(* IEC 61131-3 sources: BioPrint-Automation-Suite/projects/02_bioprint_pid/plc/src, 4 files *)

(* ---- DUT_ReferenceVectors.st ---- *)
(* =============================================================================
   DUT_ReferenceVectors — GENERATED by plc/generate_test_vectors.py. Do not edit.
   Struct types for GVL_ReferenceVectors (two DUTs in TwinCAT / CODESYS).
   ============================================================================= *)
TYPE ST_PidVector :
STRUCT
    lrSetpoint    : LREAL;
    lrMeasurement : LREAL;
    lrOutput      : LREAL;
    lrITerm       : LREAL;
END_STRUCT
END_TYPE

TYPE ST_WestgardVector :
STRUCT
    diStep     : DINT;
    lrValue    : LREAL;
    bWarn12s   : BOOL;
    bReject13s : BOOL;
    bReject22s : BOOL;
END_STRUCT
END_TYPE

(* ---- GVL_ReferenceVectors.st ---- *)
(* =============================================================================
   GVL_ReferenceVectors — GENERATED by plc/generate_test_vectors.py. Do not edit.
   Inputs and outputs of the Python reference implementation for the default
   scenario (config/default.toml), replayed scan by scan in the TcUnit tests.
   Types: DUT_ReferenceVectors.st
   ============================================================================= *)
{attribute 'qualified_only'}
VAR_GLOBAL CONSTANT
    N_VECTORS       : INT   := 300;
    LR_BASELINE_SD  : LREAL := 2.918663164239998E-01;
    aPid : ARRAY[1..300] OF ST_PidVector := [
        (lrSetpoint := 2.300000000000000E+02, lrMeasurement := 2.504570756196317E+01, lrOutput := 1.000000000000000E+02, lrITerm := 0.000000000000000E+00),
        (lrSetpoint := 2.300000000000000E+02, lrMeasurement := 2.559400238406393E+01, lrOutput := 1.000000000000000E+02, lrITerm := 0.000000000000000E+00),
        (lrSetpoint := 2.300000000000000E+02, lrMeasurement := 2.721106767937097E+01, lrOutput := 1.000000000000000E+02, lrITerm := 0.000000000000000E+00),
        (lrSetpoint := 2.300000000000000E+02, lrMeasurement := 2.906538770745868E+01, lrOutput := 1.000000000000000E+02, lrITerm := 0.000000000000000E+00),
        (lrSetpoint := 2.300000000000000E+02, lrMeasurement := 3.083779911570193E+01, lrOutput := 1.000000000000000E+02, lrITerm := 0.000000000000000E+00),
        (lrSetpoint := 2.300000000000000E+02, lrMeasurement := 3.344406655918265E+01, lrOutput := 1.000000000000000E+02, lrITerm := 0.000000000000000E+00),
        (lrSetpoint := 2.300000000000000E+02, lrMeasurement := 3.640825075871666E+01, lrOutput := 1.000000000000000E+02, lrITerm := 0.000000000000000E+00),
        (lrSetpoint := 2.300000000000000E+02, lrMeasurement := 3.928242815999355E+01, lrOutput := 1.000000000000000E+02, lrITerm := 0.000000000000000E+00),
        (lrSetpoint := 2.300000000000000E+02, lrMeasurement := 4.241953904612176E+01, lrOutput := 1.000000000000000E+02, lrITerm := 0.000000000000000E+00),
        (lrSetpoint := 2.300000000000000E+02, lrMeasurement := 4.550594203217187E+01, lrOutput := 1.000000000000000E+02, lrITerm := 0.000000000000000E+00),
        (lrSetpoint := 2.300000000000000E+02, lrMeasurement := 4.907188733629471E+01, lrOutput := 1.000000000000000E+02, lrITerm := 0.000000000000000E+00),
        (lrSetpoint := 2.300000000000000E+02, lrMeasurement := 5.243664392789950E+01, lrOutput := 1.000000000000000E+02, lrITerm := 0.000000000000000E+00),
        (lrSetpoint := 2.300000000000000E+02, lrMeasurement := 5.576754175418417E+01, lrOutput := 1.000000000000000E+02, lrITerm := 0.000000000000000E+00),
        (lrSetpoint := 2.300000000000000E+02, lrMeasurement := 5.940904962608809E+01, lrOutput := 1.000000000000000E+02, lrITerm := 0.000000000000000E+00),
        (lrSetpoint := 2.300000000000000E+02, lrMeasurement := 6.282668317532421E+01, lrOutput := 1.000000000000000E+02, lrITerm := 0.000000000000000E+00),
        (lrSetpoint := 2.300000000000000E+02, lrMeasurement := 6.617020839567282E+01, lrOutput := 1.000000000000000E+02, lrITerm := 0.000000000000000E+00),
        (lrSetpoint := 2.300000000000000E+02, lrMeasurement := 6.991626356192097E+01, lrOutput := 1.000000000000000E+02, lrITerm := 0.000000000000000E+00),
        (lrSetpoint := 2.300000000000000E+02, lrMeasurement := 7.329295415928244E+01, lrOutput := 1.000000000000000E+02, lrITerm := 0.000000000000000E+00),
        (lrSetpoint := 2.300000000000000E+02, lrMeasurement := 7.715412652709350E+01, lrOutput := 1.000000000000000E+02, lrITerm := 0.000000000000000E+00),
        (lrSetpoint := 2.300000000000000E+02, lrMeasurement := 8.060678218175724E+01, lrOutput := 1.000000000000000E+02, lrITerm := 0.000000000000000E+00),
        (lrSetpoint := 2.300000000000000E+02, lrMeasurement := 8.418207861531381E+01, lrOutput := 1.000000000000000E+02, lrITerm := 0.000000000000000E+00),
        (lrSetpoint := 2.300000000000000E+02, lrMeasurement := 8.770466127710711E+01, lrOutput := 1.000000000000000E+02, lrITerm := 0.000000000000000E+00),
        (lrSetpoint := 2.300000000000000E+02, lrMeasurement := 9.158689819204071E+01, lrOutput := 1.000000000000000E+02, lrITerm := 0.000000000000000E+00),
        (lrSetpoint := 2.300000000000000E+02, lrMeasurement := 9.497539444205835E+01, lrOutput := 1.000000000000000E+02, lrITerm := 0.000000000000000E+00),
        (lrSetpoint := 2.300000000000000E+02, lrMeasurement := 9.852661866900469E+01, lrOutput := 1.000000000000000E+02, lrITerm := 0.000000000000000E+00),
        (lrSetpoint := 2.300000000000000E+02, lrMeasurement := 1.021266989746227E+02, lrOutput := 1.000000000000000E+02, lrITerm := 0.000000000000000E+00),
        (lrSetpoint := 2.300000000000000E+02, lrMeasurement := 1.058436726674556E+02, lrOutput := 1.000000000000000E+02, lrITerm := 0.000000000000000E+00),
        (lrSetpoint := 2.300000000000000E+02, lrMeasurement := 1.093980483030509E+02, lrOutput := 1.000000000000000E+02, lrITerm := 0.000000000000000E+00),
        (lrSetpoint := 2.300000000000000E+02, lrMeasurement := 1.129792015668312E+02, lrOutput := 1.000000000000000E+02, lrITerm := 0.000000000000000E+00),
        (lrSetpoint := 2.300000000000000E+02, lrMeasurement := 1.165502773982586E+02, lrOutput := 1.000000000000000E+02, lrITerm := 0.000000000000000E+00),
        (lrSetpoint := 2.300000000000000E+02, lrMeasurement := 1.203692878042951E+02, lrOutput := 1.000000000000000E+02, lrITerm := 0.000000000000000E+00),
        (lrSetpoint := 2.300000000000000E+02, lrMeasurement := 1.235432685102606E+02, lrOutput := 1.000000000000000E+02, lrITerm := 0.000000000000000E+00),
        (lrSetpoint := 2.300000000000000E+02, lrMeasurement := 1.270772148357379E+02, lrOutput := 1.000000000000000E+02, lrITerm := 0.000000000000000E+00),
        (lrSetpoint := 2.300000000000000E+02, lrMeasurement := 1.305753003884958E+02, lrOutput := 1.000000000000000E+02, lrITerm := 0.000000000000000E+00),
        (lrSetpoint := 2.300000000000000E+02, lrMeasurement := 1.343264670026235E+02, lrOutput := 1.000000000000000E+02, lrITerm := 0.000000000000000E+00),
        (lrSetpoint := 2.300000000000000E+02, lrMeasurement := 1.379334266122466E+02, lrOutput := 1.000000000000000E+02, lrITerm := 0.000000000000000E+00),
        (lrSetpoint := 2.300000000000000E+02, lrMeasurement := 1.412702435435773E+02, lrOutput := 1.000000000000000E+02, lrITerm := 0.000000000000000E+00),
        (lrSetpoint := 2.300000000000000E+02, lrMeasurement := 1.446777639636957E+02, lrOutput := 1.000000000000000E+02, lrITerm := 0.000000000000000E+00),
        (lrSetpoint := 2.300000000000000E+02, lrMeasurement := 1.481897288334872E+02, lrOutput := 1.000000000000000E+02, lrITerm := 0.000000000000000E+00),
        (lrSetpoint := 2.300000000000000E+02, lrMeasurement := 1.519137400563598E+02, lrOutput := 1.000000000000000E+02, lrITerm := 0.000000000000000E+00),
        (lrSetpoint := 2.300000000000000E+02, lrMeasurement := 1.554235085010919E+02, lrOutput := 1.000000000000000E+02, lrITerm := 0.000000000000000E+00),
        (lrSetpoint := 2.300000000000000E+02, lrMeasurement := 1.588824707065076E+02, lrOutput := 1.000000000000000E+02, lrITerm := 0.000000000000000E+00),
        (lrSetpoint := 2.300000000000000E+02, lrMeasurement := 1.621832501003170E+02, lrOutput := 1.000000000000000E+02, lrITerm := 0.000000000000000E+00),
        (lrSetpoint := 2.300000000000000E+02, lrMeasurement := 1.657930793899823E+02, lrOutput := 1.000000000000000E+02, lrITerm := 0.000000000000000E+00),
        (lrSetpoint := 2.300000000000000E+02, lrMeasurement := 1.692440373830902E+02, lrOutput := 1.000000000000000E+02, lrITerm := 0.000000000000000E+00),
        (lrSetpoint := 2.300000000000000E+02, lrMeasurement := 1.727207213966689E+02, lrOutput := 1.000000000000000E+02, lrITerm := 0.000000000000000E+00),
        (lrSetpoint := 2.300000000000000E+02, lrMeasurement := 1.762731259192086E+02, lrOutput := 1.000000000000000E+02, lrITerm := 0.000000000000000E+00),
        (lrSetpoint := 2.300000000000000E+02, lrMeasurement := 1.796235615768844E+02, lrOutput := 1.000000000000000E+02, lrITerm := 0.000000000000000E+00),
        (lrSetpoint := 2.300000000000000E+02, lrMeasurement := 1.831325956067453E+02, lrOutput := 1.000000000000000E+02, lrITerm := 0.000000000000000E+00),
        (lrSetpoint := 2.300000000000000E+02, lrMeasurement := 1.864747670133277E+02, lrOutput := 1.000000000000000E+02, lrITerm := 0.000000000000000E+00),
        (lrSetpoint := 2.300000000000000E+02, lrMeasurement := 1.899350152806136E+02, lrOutput := 1.000000000000000E+02, lrITerm := 0.000000000000000E+00),
        (lrSetpoint := 2.300000000000000E+02, lrMeasurement := 1.934065144925135E+02, lrOutput := 1.000000000000000E+02, lrITerm := 0.000000000000000E+00),
        (lrSetpoint := 2.300000000000000E+02, lrMeasurement := 1.965065899891975E+02, lrOutput := 1.000000000000000E+02, lrITerm := 0.000000000000000E+00),
        (lrSetpoint := 2.300000000000000E+02, lrMeasurement := 2.000837349498422E+02, lrOutput := 1.000000000000000E+02, lrITerm := 0.000000000000000E+00),
        (lrSetpoint := 2.300000000000000E+02, lrMeasurement := 2.034608444403627E+02, lrOutput := 1.000000000000000E+02, lrITerm := 0.000000000000000E+00),
        (lrSetpoint := 2.300000000000000E+02, lrMeasurement := 2.068284883225735E+02, lrOutput := 1.000000000000000E+02, lrITerm := 0.000000000000000E+00),
        (lrSetpoint := 2.300000000000000E+02, lrMeasurement := 2.102691859917106E+02, lrOutput := 9.423082560990316E+01, lrITerm := 4.932703502072343E+00),
        (lrSetpoint := 2.300000000000000E+02, lrMeasurement := 2.138707975791627E+02, lrOutput := 6.666316008304979E+01, lrITerm := 8.965004107281665E+00),
        (lrSetpoint := 2.300000000000000E+02, lrMeasurement := 2.166047382771748E+02, lrOutput := 6.146576947420901E+01, lrITerm := 1.231381953798795E+01),
        (lrSetpoint := 2.300000000000000E+02, lrMeasurement := 2.196531259180408E+02, lrOutput := 3.729929969102109E+01, lrITerm := 1.490053805847776E+01),
        (lrSetpoint := 2.300000000000000E+02, lrMeasurement := 2.215944746720401E+02, lrOutput := 4.110929574553012E+01, lrITerm := 1.700191939046773E+01),
        (lrSetpoint := 2.300000000000000E+02, lrMeasurement := 2.238164015632227E+02, lrOutput := 2.383841098123746E+01, lrITerm := 1.854781899966206E+01),
        (lrSetpoint := 2.300000000000000E+02, lrMeasurement := 2.255252359017419E+02, lrOutput := 1.928763429145494E+01, lrITerm := 1.966651002422659E+01),
        (lrSetpoint := 2.300000000000000E+02, lrMeasurement := 2.268803103257552E+02, lrOutput := 1.648736134876521E+01, lrITerm := 2.044643244278778E+01),
        (lrSetpoint := 2.300000000000000E+02, lrMeasurement := 2.278955664907341E+02, lrOutput := 1.578059255697349E+01, lrITerm := 2.097254082010426E+01),
        (lrSetpoint := 2.300000000000000E+02, lrMeasurement := 2.286631929043172E+02, lrOutput := 1.531369347470648E+01, lrITerm := 2.130674259402496E+01),
        (lrSetpoint := 2.300000000000000E+02, lrMeasurement := 2.290508932078158E+02, lrOutput := 1.959616759661151E+01, lrITerm := 2.154401929207102E+01),
        (lrSetpoint := 2.300000000000000E+02, lrMeasurement := 2.294681164603311E+02, lrOutput := 1.734834524750830E+01, lrITerm := 2.167699017698826E+01),
        (lrSetpoint := 2.300000000000000E+02, lrMeasurement := 2.299838292420773E+02, lrOutput := 1.184225177254323E+01, lrITerm := 2.168103286646892E+01),
        (lrSetpoint := 2.300000000000000E+02, lrMeasurement := 2.300096375187556E+02, lrOutput := 1.919496147842190E+01, lrITerm := 2.167862348678002E+01),
        (lrSetpoint := 2.300000000000000E+02, lrMeasurement := 2.299780300469962E+02, lrOutput := 2.188428277554846E+01, lrITerm := 2.168411597503096E+01),
        (lrSetpoint := 2.300000000000000E+02, lrMeasurement := 2.301089493703319E+02, lrOutput := 1.869545593171979E+01, lrITerm := 2.165687863244799E+01),
        (lrSetpoint := 2.300000000000000E+02, lrMeasurement := 2.302094572798513E+02, lrOutput := 1.790276397374864E+01, lrITerm := 2.160451431248516E+01),
        (lrSetpoint := 2.300000000000000E+02, lrMeasurement := 2.304978744922259E+02, lrOutput := 1.247715593364422E+01, lrITerm := 2.148004568942869E+01),
        (lrSetpoint := 2.300000000000000E+02, lrMeasurement := 2.304858332660471E+02, lrOutput := 1.666060209980525E+01, lrITerm := 2.135858737291692E+01),
        (lrSetpoint := 2.300000000000000E+02, lrMeasurement := 2.306128359144820E+02, lrOutput := 1.410838487453493E+01, lrITerm := 2.120537839429642E+01),
        (lrSetpoint := 2.300000000000000E+02, lrMeasurement := 2.304736944247048E+02, lrOutput := 1.908480198613638E+01, lrITerm := 2.108695478812023E+01),
        (lrSetpoint := 2.300000000000000E+02, lrMeasurement := 2.306144061359000E+02, lrOutput := 1.412419730695324E+01, lrITerm := 2.093335325414524E+01),
        (lrSetpoint := 2.300000000000000E+02, lrMeasurement := 2.307194784114588E+02, lrOutput := 1.293771857867122E+01, lrITerm := 2.075348365128055E+01),
        (lrSetpoint := 2.300000000000000E+02, lrMeasurement := 2.305911113626528E+02, lrOutput := 1.751870013410300E+01, lrITerm := 2.060570581061735E+01),
        (lrSetpoint := 2.300000000000000E+02, lrMeasurement := 2.307337919192282E+02, lrOutput := 1.259741061672039E+01, lrITerm := 2.042225783081031E+01),
        (lrSetpoint := 2.300000000000000E+02, lrMeasurement := 2.305232005023320E+02, lrOutput := 1.908441398485769E+01, lrITerm := 2.029145770522732E+01),
        (lrSetpoint := 2.300000000000000E+02, lrMeasurement := 2.305177106373760E+02, lrOutput := 1.670389484582921E+01, lrITerm := 2.016203004588333E+01),
        (lrSetpoint := 2.300000000000000E+02, lrMeasurement := 2.304407682616513E+02, lrOutput := 1.789347987864461E+01, lrITerm := 2.005183798047049E+01),
        (lrSetpoint := 2.300000000000000E+02, lrMeasurement := 2.302345111439646E+02, lrOutput := 2.169079252402655E+01, lrITerm := 1.999321019447934E+01),
        (lrSetpoint := 2.300000000000000E+02, lrMeasurement := 2.304233655001475E+02, lrOutput := 1.419350941559006E+01, lrITerm := 1.988736881944247E+01),
        (lrSetpoint := 2.300000000000000E+02, lrMeasurement := 2.301765571888204E+02, lrOutput := 2.191831791237351E+01, lrITerm := 1.984322952223738E+01),
        (lrSetpoint := 2.300000000000000E+02, lrMeasurement := 2.301718013630896E+02, lrOutput := 1.919947066857960E+01, lrITerm := 1.980027918146497E+01),
        (lrSetpoint := 2.300000000000000E+02, lrMeasurement := 2.301656351697725E+02, lrOutput := 1.868716860228188E+01, lrITerm := 1.975887038902184E+01),
        (lrSetpoint := 2.300000000000000E+02, lrMeasurement := 2.300808227245562E+02, lrOutput := 2.049975794918330E+01, lrITerm := 1.973866470788280E+01),
        (lrSetpoint := 2.300000000000000E+02, lrMeasurement := 2.300450161809068E+02, lrOutput := 2.022172092134138E+01, lrITerm := 1.972741066265610E+01),
        (lrSetpoint := 2.300000000000000E+02, lrMeasurement := 2.298685710227648E+02, lrOutput := 2.380571019630718E+01, lrITerm := 1.976026790696491E+01),
        (lrSetpoint := 2.300000000000000E+02, lrMeasurement := 2.297903074584952E+02, lrOutput := 2.334125049698557E+01, lrITerm := 1.981269104234112E+01),
        (lrSetpoint := 2.300000000000000E+02, lrMeasurement := 2.298346004226570E+02, lrOutput := 2.083875395335288E+01, lrITerm := 1.985404093667687E+01),
        (lrSetpoint := 2.300000000000000E+02, lrMeasurement := 2.295852197770309E+02, lrOutput := 2.719837138577611E+01, lrITerm := 1.995773599241915E+01),
        (lrSetpoint := 2.300000000000000E+02, lrMeasurement := 2.296599261274224E+02, lrOutput := 2.235252255684210E+01, lrITerm := 2.004275446056356E+01),
        (lrSetpoint := 2.300000000000000E+02, lrMeasurement := 2.297182708644902E+02, lrOutput := 2.135133945856617E+01, lrITerm := 2.011318674444102E+01),
        (lrSetpoint := 2.300000000000000E+02, lrMeasurement := 2.298000366341335E+02, lrOutput := 2.025149612455615E+01, lrITerm := 2.016317758590765E+01),
        (lrSetpoint := 2.300000000000000E+02, lrMeasurement := 2.300288961980845E+02, lrOutput := 1.596075325083648E+01, lrITerm := 2.015595353638652E+01),
        (lrSetpoint := 2.300000000000000E+02, lrMeasurement := 2.298093482091375E+02, lrOutput := 2.444879249397976E+01, lrITerm := 2.020361648410214E+01),
        (lrSetpoint := 2.300000000000000E+02, lrMeasurement := 2.298940447799201E+02, lrOutput := 2.026659425383454E+01, lrITerm := 2.023010528912211E+01),
        (lrSetpoint := 2.300000000000000E+02, lrMeasurement := 2.301432779377677E+02, lrOutput := 1.489810121779246E+01, lrITerm := 2.019428580468018E+01),
        (lrSetpoint := 2.300000000000000E+02, lrMeasurement := 2.298459618394776E+02, lrOutput := 2.539216598468198E+01, lrITerm := 2.023279534481078E+01),
        (lrSetpoint := 2.300000000000000E+02, lrMeasurement := 2.300026310488091E+02, lrOutput := 1.848979491396977E+01, lrITerm := 2.023213758260850E+01),
        (lrSetpoint := 2.300000000000000E+02, lrMeasurement := 2.297259479761731E+02, lrOutput := 2.657573708572423E+01, lrITerm := 2.030065058856523E+01),
        (lrSetpoint := 2.300000000000000E+02, lrMeasurement := 2.298549920521735E+02, lrOutput := 2.024879500343473E+01, lrITerm := 2.033690257552185E+01),
        (lrSetpoint := 2.300000000000000E+02, lrMeasurement := 2.297521760524508E+02, lrOutput := 2.377687190742672E+01, lrITerm := 2.039885856240915E+01),
        (lrSetpoint := 2.300000000000000E+02, lrMeasurement := 2.298704273997785E+02, lrOutput := 1.985489530991842E+01, lrITerm := 2.043125171246452E+01),
        (lrSetpoint := 2.300000000000000E+02, lrMeasurement := 2.300586262338561E+02, lrOutput := 1.661381649704559E+01, lrITerm := 2.041659515400049E+01),
        (lrSetpoint := 2.300000000000000E+02, lrMeasurement := 2.296482659229140E+02, lrOutput := 2.921741250781378E+01, lrITerm := 2.050452867327200E+01),
        (lrSetpoint := 2.300000000000000E+02, lrMeasurement := 2.300127602678513E+02, lrOutput := 1.574714918807162E+01, lrITerm := 2.050133860630917E+01),
        (lrSetpoint := 2.300000000000000E+02, lrMeasurement := 2.299745877595838E+02, lrOutput := 2.039132826693744E+01, lrITerm := 2.050769166641322E+01),
        (lrSetpoint := 2.300000000000000E+02, lrMeasurement := 2.298370036522997E+02, lrOutput := 2.398982498692613E+01, lrITerm := 2.054844075333830E+01),
        (lrSetpoint := 2.300000000000000E+02, lrMeasurement := 2.297662189294558E+02, lrOutput := 2.403717284122651E+01, lrITerm := 2.060688602097434E+01),
        (lrSetpoint := 2.300000000000000E+02, lrMeasurement := 2.301069608762478E+02, lrOutput := 1.458459529443878E+01, lrITerm := 2.058014580191240E+01),
        (lrSetpoint := 2.300000000000000E+02, lrMeasurement := 2.301034615741697E+02, lrOutput := 1.875460394876319E+01, lrITerm := 2.055428040836998E+01),
        (lrSetpoint := 2.300000000000000E+02, lrMeasurement := 2.303148002423178E+02, lrOutput := 1.438136294562796E+01, lrITerm := 2.047558034779052E+01),
        (lrSetpoint := 2.300000000000000E+02, lrMeasurement := 2.303555301449315E+02, lrOutput := 1.617561511756174E+01, lrITerm := 2.038669781155763E+01),
        (lrSetpoint := 2.300000000000000E+02, lrMeasurement := 2.306586161636685E+02, lrOutput := 9.830369854592995E+00, lrITerm := 2.022204377064051E+01),
        (lrSetpoint := 2.300000000000000E+02, lrMeasurement := 2.303959258597061E+02, lrOutput := 2.013415137012417E+01, lrITerm := 2.012306230571399E+01),
        (lrSetpoint := 2.300000000000000E+02, lrMeasurement := 2.303270774525105E+02, lrOutput := 1.916194702604438E+01, lrITerm := 2.004129294258638E+01),
        (lrSetpoint := 2.300000000000000E+02, lrMeasurement := 2.305308276598897E+02, lrOutput := 1.274941617113750E+01, lrITerm := 1.990858602761396E+01),
        (lrSetpoint := 2.300000000000000E+02, lrMeasurement := 2.304918859423371E+02, lrOutput := 1.589108476870233E+01, lrITerm := 1.978561454202969E+01),
        (lrSetpoint := 2.300000000000000E+02, lrMeasurement := 2.305868168294902E+02, lrOutput := 1.343359305736029E+01, lrITerm := 1.963891033465715E+01),
        (lrSetpoint := 2.300000000000000E+02, lrMeasurement := 2.303892627913187E+02, lrOutput := 1.928620038874604E+01, lrITerm := 1.954159463682747E+01),
        (lrSetpoint := 2.300000000000000E+02, lrMeasurement := 2.302083083202458E+02, lrOutput := 2.129006414846046E+01, lrITerm := 1.948951755676602E+01),
        (lrSetpoint := 2.300000000000000E+02, lrMeasurement := 2.302879174462091E+02, lrOutput := 1.653385524086008E+01, lrITerm := 1.941753819521375E+01),
        (lrSetpoint := 2.300000000000000E+02, lrMeasurement := 2.297863666250582E+02, lrOutput := 2.908875799996291E+01, lrITerm := 1.947094653894921E+01),
        (lrSetpoint := 2.300000000000000E+02, lrMeasurement := 2.298453652638796E+02, lrOutput := 2.138445378309544E+01, lrITerm := 1.950960522297932E+01),
        (lrSetpoint := 2.300000000000000E+02, lrMeasurement := 2.297852853998048E+02, lrOutput := 2.236983263401705E+01, lrITerm := 1.956328387302812E+01),
        (lrSetpoint := 2.300000000000000E+02, lrMeasurement := 2.298611656666668E+02, lrOutput := 1.971234924511949E+01, lrITerm := 1.959799245636141E+01),
        (lrSetpoint := 2.300000000000000E+02, lrMeasurement := 2.296984707598905E+02, lrOutput := 2.448946362010373E+01, lrITerm := 1.967337476638878E+01),
        (lrSetpoint := 2.300000000000000E+02, lrMeasurement := 2.300134306392112E+02, lrOutput := 1.500398491033279E+01, lrITerm := 1.967001710658597E+01),
        (lrSetpoint := 2.300000000000000E+02, lrMeasurement := 2.298490494877590E+02, lrOutput := 2.263373983929725E+01, lrITerm := 1.970775473464622E+01),
        (lrSetpoint := 2.300000000000000E+02, lrMeasurement := 2.296442219691345E+02, lrOutput := 2.626383998862416E+01, lrITerm := 1.979669924236260E+01),
        (lrSetpoint := 2.300000000000000E+02, lrMeasurement := 2.297367369885094E+02, lrOutput := 2.121256207702870E+01, lrITerm := 1.986251499523525E+01),
        (lrSetpoint := 2.300000000000000E+02, lrMeasurement := 2.299557157451501E+02, lrOutput := 1.657298858946894E+01, lrITerm := 1.987358605894772E+01),
        (lrSetpoint := 2.300000000000000E+02, lrMeasurement := 2.300155318818599E+02, lrOutput := 1.805741554459039E+01, lrITerm := 1.986970308848274E+01),
        (lrSetpoint := 2.300000000000000E+02, lrMeasurement := 2.301509214398248E+02, lrOutput := 1.612076178468788E+01, lrITerm := 1.983197272852654E+01),
        (lrSetpoint := 2.300000000000000E+02, lrMeasurement := 2.302200352161047E+02, lrOutput := 1.641009389013652E+01, lrITerm := 1.977696392450036E+01),
        (lrSetpoint := 2.300000000000000E+02, lrMeasurement := 2.297549336201718E+02, lrOutput := 2.891906943190371E+01, lrITerm := 1.983823051945741E+01),
        (lrSetpoint := 2.300000000000000E+02, lrMeasurement := 2.295307302659245E+02, lrOutput := 2.872102106830100E+01, lrITerm := 1.995554795297628E+01),
        (lrSetpoint := 2.300000000000000E+02, lrMeasurement := 2.294052885678543E+02, lrOutput := 2.787124748584564E+01, lrITerm := 2.010422581101270E+01),
        (lrSetpoint := 2.300000000000000E+02, lrMeasurement := 2.298522298602363E+02, lrOutput := 1.477413482948581E+01, lrITerm := 2.014116834595364E+01),
        (lrSetpoint := 2.300000000000000E+02, lrMeasurement := 2.297115211052058E+02, lrOutput := 2.346262038157825E+01, lrITerm := 2.021328806965219E+01),
        (lrSetpoint := 2.300000000000000E+02, lrMeasurement := 2.298054273966737E+02, lrOutput := 2.050431161432098E+01, lrITerm := 2.026193122048376E+01),
        (lrSetpoint := 2.300000000000000E+02, lrMeasurement := 2.297982350513737E+02, lrOutput := 2.177872948489685E+01, lrITerm := 2.031237245764034E+01),
        (lrSetpoint := 2.300000000000000E+02, lrMeasurement := 2.298912673017996E+02, lrOutput := 1.969134869862730E+01, lrITerm := 2.033955563219043E+01),
        (lrSetpoint := 2.300000000000000E+02, lrMeasurement := 2.300789608336171E+02, lrOutput := 1.638141854193576E+01, lrITerm := 2.031981542378614E+01),
        (lrSetpoint := 2.300000000000000E+02, lrMeasurement := 2.299119910387465E+02, lrOutput := 2.305606402947607E+01, lrITerm := 2.034181766409952E+01),
        (lrSetpoint := 2.300000000000000E+02, lrMeasurement := 2.298543613889811E+02, lrOutput := 2.286744553632186E+01, lrITerm := 2.037822731685426E+01),
        (lrSetpoint := 2.300000000000000E+02, lrMeasurement := 2.294720232167521E+02, lrOutput := 3.111626840057623E+01, lrITerm := 2.051022151266623E+01),
        (lrSetpoint := 2.300000000000000E+02, lrMeasurement := 2.289971171519480E+02, lrOutput := 3.765894857034665E+01, lrITerm := 2.076094222467924E+01),
        (lrSetpoint := 2.300000000000000E+02, lrMeasurement := 2.287900661865506E+02, lrOutput := 3.583070034424563E+01, lrITerm := 2.106342567804160E+01),
        (lrSetpoint := 2.300000000000000E+02, lrMeasurement := 2.284515985235186E+02, lrOutput := 4.027078129924619E+01, lrITerm := 2.145052604716194E+01),
        (lrSetpoint := 2.300000000000000E+02, lrMeasurement := 2.283411627174421E+02, lrOutput := 3.818951521353537E+01, lrITerm := 2.186523536780142E+01),
        (lrSetpoint := 2.300000000000000E+02, lrMeasurement := 2.277124386479682E+02, lrOutput := 5.140791795070005E+01, lrITerm := 2.243712570580936E+01),
        (lrSetpoint := 2.300000000000000E+02, lrMeasurement := 2.275574921917000E+02, lrOutput := 4.720101871030254E+01, lrITerm := 2.304775265788436E+01),
        (lrSetpoint := 2.300000000000000E+02, lrMeasurement := 2.271008315546960E+02, lrOutput := 5.519510324090932E+01, lrITerm := 2.377254476921035E+01),
        (lrSetpoint := 2.300000000000000E+02, lrMeasurement := 2.268624201050854E+02, lrOutput := 5.511800427788045E+01, lrITerm := 2.455693974293901E+01),
        (lrSetpoint := 2.300000000000000E+02, lrMeasurement := 2.268378562653796E+02, lrOutput := 5.212973206397371E+01, lrITerm := 2.534747567659410E+01),
        (lrSetpoint := 2.300000000000000E+02, lrMeasurement := 2.268104966628377E+02, lrOutput := 5.239565315093742E+01, lrITerm := 2.614485151088468E+01),
        (lrSetpoint := 2.300000000000000E+02, lrMeasurement := 2.271727202882387E+02, lrOutput := 4.382128611504928E+01, lrITerm := 2.685167143882499E+01),
        (lrSetpoint := 2.300000000000000E+02, lrMeasurement := 2.265982553891899E+02, lrOutput := 6.297777825921683E+01, lrITerm := 2.770210759152752E+01),
        (lrSetpoint := 2.300000000000000E+02, lrMeasurement := 2.268067431131597E+02, lrOutput := 5.232301608068577E+01, lrITerm := 2.850042181323761E+01),
        (lrSetpoint := 2.300000000000000E+02, lrMeasurement := 2.264977102339018E+02, lrOutput := 6.199414628621889E+01, lrITerm := 2.937599425476216E+01),
        (lrSetpoint := 2.300000000000000E+02, lrMeasurement := 2.267918815203126E+02, lrOutput := 5.205619791014471E+01, lrITerm := 3.017802387468402E+01),
        (lrSetpoint := 2.300000000000000E+02, lrMeasurement := 2.267072664589627E+02, lrOutput := 5.793956180943100E+01, lrITerm := 3.100120725994333E+01),
        (lrSetpoint := 2.300000000000000E+02, lrMeasurement := 2.266504042455074E+02, lrOutput := 5.966446489403108E+01, lrITerm := 3.183860619856648E+01),
        (lrSetpoint := 2.300000000000000E+02, lrMeasurement := 2.267264485475885E+02, lrOutput := 5.783451537956719E+01, lrITerm := 3.265699406166934E+01),
        (lrSetpoint := 2.300000000000000E+02, lrMeasurement := 2.267063455066636E+02, lrOutput := 5.994911422621549E+01, lrITerm := 3.348040768500345E+01),
        (lrSetpoint := 2.300000000000000E+02, lrMeasurement := 2.269697698730993E+02, lrOutput := 5.428891048786628E+01, lrITerm := 3.423796521672862E+01),
        (lrSetpoint := 2.300000000000000E+02, lrMeasurement := 2.269111095789345E+02, lrOutput := 5.982169674834228E+01, lrITerm := 3.501018782199499E+01),
        (lrSetpoint := 2.300000000000000E+02, lrMeasurement := 2.268960923785198E+02, lrOutput := 6.087777801740615E+01, lrITerm := 3.578616472736503E+01),
        (lrSetpoint := 2.300000000000000E+02, lrMeasurement := 2.270156326598504E+02, lrOutput := 5.854662124594902E+01, lrITerm := 3.653225656240242E+01),
        (lrSetpoint := 2.300000000000000E+02, lrMeasurement := 2.273641290287552E+02, lrOutput := 5.233013536516516E+01, lrITerm := 3.719122430521362E+01),
        (lrSetpoint := 2.300000000000000E+02, lrMeasurement := 2.276619484977107E+02, lrOutput := 5.052542635381054E+01, lrITerm := 3.777573718078593E+01),
        (lrSetpoint := 2.300000000000000E+02, lrMeasurement := 2.274873010596821E+02, lrOutput := 6.010891787780903E+01, lrITerm := 3.840391191586541E+01),
        (lrSetpoint := 2.300000000000000E+02, lrMeasurement := 2.275169921363721E+02, lrOutput := 5.873435245163500E+01, lrITerm := 3.902466388177238E+01),
        (lrSetpoint := 2.300000000000000E+02, lrMeasurement := 2.276650690346880E+02, lrOutput := 5.588773910470954E+01, lrITerm := 3.960839662310037E+01),
        (lrSetpoint := 2.300000000000000E+02, lrMeasurement := 2.278966070310045E+02, lrOutput := 5.277675962807260E+01, lrITerm := 4.013424486534925E+01),
        (lrSetpoint := 2.300000000000000E+02, lrMeasurement := 2.277815965043510E+02, lrOutput := 5.943931633306123E+01, lrITerm := 4.068884573926150E+01),
        (lrSetpoint := 2.300000000000000E+02, lrMeasurement := 2.277607171447250E+02, lrOutput := 5.969764757501729E+01, lrITerm := 4.124866645308024E+01),
        (lrSetpoint := 2.300000000000000E+02, lrMeasurement := 2.280841211516531E+02, lrOutput := 5.198714649704154E+01, lrITerm := 4.172763616516698E+01),
        (lrSetpoint := 2.300000000000000E+02, lrMeasurement := 2.280378619566982E+02, lrOutput := 5.764191805070404E+01, lrITerm := 4.221817067599243E+01),
        (lrSetpoint := 2.300000000000000E+02, lrMeasurement := 2.282695321084727E+02, lrOutput := 5.273313695836017E+01, lrITerm := 4.265078764887425E+01),
        (lrSetpoint := 2.300000000000000E+02, lrMeasurement := 2.281034579844685E+02, lrOutput := 6.020216649652940E+01, lrITerm := 4.312492315275712E+01),
        (lrSetpoint := 2.300000000000000E+02, lrMeasurement := 2.279622185203662E+02, lrOutput := 6.257743322927701E+01, lrITerm := 4.363436852266557E+01),
        (lrSetpoint := 2.300000000000000E+02, lrMeasurement := 2.280545056773856E+02, lrOutput := 5.873626474583284E+01, lrITerm := 4.412074210331917E+01),
        (lrSetpoint := 2.300000000000000E+02, lrMeasurement := 2.286269974803834E+02, lrOutput := 4.609845765451041E+01, lrITerm := 4.446399273322332E+01),
        (lrSetpoint := 2.300000000000000E+02, lrMeasurement := 2.286671160554017E+02, lrOutput := 5.294847702873701E+01, lrITerm := 4.479721371937289E+01),
        (lrSetpoint := 2.300000000000000E+02, lrMeasurement := 2.283905080974753E+02, lrOutput := 6.199888759253917E+01, lrITerm := 4.519958669500406E+01),
        (lrSetpoint := 2.300000000000000E+02, lrMeasurement := 2.284205711481603E+02, lrOutput := 5.853353904719056E+01, lrITerm := 4.559444390796399E+01),
        (lrSetpoint := 2.300000000000000E+02, lrMeasurement := 2.288186192176935E+02, lrOutput := 4.903279911436165E+01, lrITerm := 4.588978910354061E+01),
        (lrSetpoint := 2.300000000000000E+02, lrMeasurement := 2.285314344307211E+02, lrOutput := 6.133880439212427E+01, lrITerm := 4.625693049586033E+01),
        (lrSetpoint := 2.300000000000000E+02, lrMeasurement := 2.287350459843640E+02, lrOutput := 5.410168613497742E+01, lrITerm := 4.657316899976933E+01),
        (lrSetpoint := 2.300000000000000E+02, lrMeasurement := 2.291414097941779E+02, lrOutput := 4.663649424280365E+01, lrITerm := 4.678781655122486E+01),
        (lrSetpoint := 2.300000000000000E+02, lrMeasurement := 2.291081848729324E+02, lrOutput := 5.327288129846185E+01, lrITerm := 4.701077033299177E+01),
        (lrSetpoint := 2.300000000000000E+02, lrMeasurement := 2.292964414262748E+02, lrOutput := 4.962854170253177E+01, lrITerm := 4.718665997642307E+01),
        (lrSetpoint := 2.300000000000000E+02, lrMeasurement := 2.293808272853664E+02, lrOutput := 5.030734375394525E+01, lrITerm := 4.734145315508147E+01),
        (lrSetpoint := 2.300000000000000E+02, lrMeasurement := 2.295518096900797E+02, lrOutput := 4.790580651287138E+01, lrITerm := 4.745350073256155E+01),
        (lrSetpoint := 2.300000000000000E+02, lrMeasurement := 2.297340947421611E+02, lrOutput := 4.610401493661986E+01, lrITerm := 4.751997704702129E+01),
        (lrSetpoint := 2.300000000000000E+02, lrMeasurement := 2.294861354096551E+02, lrOutput := 5.501806840283870E+01, lrITerm := 4.764844319460750E+01),
        (lrSetpoint := 2.300000000000000E+02, lrMeasurement := 2.295284263331895E+02, lrOutput := 5.151401286633974E+01, lrITerm := 4.776633661131014E+01),
        (lrSetpoint := 2.300000000000000E+02, lrMeasurement := 2.290650907176098E+02, lrOutput := 6.288772542441307E+01, lrITerm := 4.800006393190769E+01),
        (lrSetpoint := 2.300000000000000E+02, lrMeasurement := 2.293768370143731E+02, lrOutput := 4.963489526179389E+01, lrITerm := 4.815585467831442E+01),
        (lrSetpoint := 2.300000000000000E+02, lrMeasurement := 2.292258378088339E+02, lrOutput := 5.625742738375546E+01, lrITerm := 4.834939522610595E+01),
        (lrSetpoint := 2.300000000000000E+02, lrMeasurement := 2.291530512192492E+02, lrOutput := 5.684425502631954E+01, lrITerm := 4.856113242129366E+01),
        (lrSetpoint := 2.300000000000000E+02, lrMeasurement := 2.292043165056924E+02, lrOutput := 5.460678313804437E+01, lrITerm := 4.876005329487057E+01),
        (lrSetpoint := 2.300000000000000E+02, lrMeasurement := 2.292824733439275E+02, lrOutput := 5.332539117344817E+01, lrITerm := 4.893943495888869E+01),
        (lrSetpoint := 2.300000000000000E+02, lrMeasurement := 2.294540619211454E+02, lrOutput := 5.042715546714970E+01, lrITerm := 4.907591947860234E+01),
        (lrSetpoint := 2.300000000000000E+02, lrMeasurement := 2.290702146383318E+02, lrOutput := 6.228495150892357E+01, lrITerm := 4.930836581901939E+01),
        (lrSetpoint := 2.300000000000000E+02, lrMeasurement := 2.292902545832142E+02, lrOutput := 5.275078694869494E+01, lrITerm := 4.948580217321582E+01),
        (lrSetpoint := 2.300000000000000E+02, lrMeasurement := 2.292086951375199E+02, lrOutput := 5.683642270802495E+01, lrITerm := 4.968362838883585E+01),
        (lrSetpoint := 2.300000000000000E+02, lrMeasurement := 2.292419763819967E+02, lrOutput := 5.556929440960266E+01, lrITerm := 4.987313429333666E+01),
        (lrSetpoint := 2.300000000000000E+02, lrMeasurement := 2.294530367481974E+02, lrOutput := 5.093500949594558E+01, lrITerm := 5.000987510628731E+01),
        (lrSetpoint := 2.300000000000000E+02, lrMeasurement := 2.293613959075460E+02, lrOutput := 5.605449799450183E+01, lrITerm := 5.016952612940080E+01),
        (lrSetpoint := 2.300000000000000E+02, lrMeasurement := 2.294712797684037E+02, lrOutput := 5.292855409144251E+01, lrITerm := 5.030170618729989E+01),
        (lrSetpoint := 2.300000000000000E+02, lrMeasurement := 2.292235190820188E+02, lrOutput := 6.035126195307738E+01, lrITerm := 5.049582641679519E+01),
        (lrSetpoint := 2.300000000000000E+02, lrMeasurement := 2.291629751724858E+02, lrOutput := 5.909870143480222E+01, lrITerm := 5.070508262367375E+01),
        (lrSetpoint := 2.300000000000000E+02, lrMeasurement := 2.292804089571940E+02, lrOutput := 5.510225220969527E+01, lrITerm := 5.088498038437525E+01),
        (lrSetpoint := 2.300000000000000E+02, lrMeasurement := 2.293874877761780E+02, lrOutput := 5.391705382373650E+01, lrITerm := 5.103810844033075E+01),
        (lrSetpoint := 2.300000000000000E+02, lrMeasurement := 2.293982407687014E+02, lrOutput := 5.542634373673484E+01, lrITerm := 5.118854824815539E+01),
        (lrSetpoint := 2.300000000000000E+02, lrMeasurement := 2.292279554865906E+02, lrOutput := 6.016722432519352E+01, lrITerm := 5.138155937650773E+01),
        (lrSetpoint := 2.300000000000000E+02, lrMeasurement := 2.294571546504262E+02, lrOutput := 5.271470865740443E+01, lrITerm := 5.151727071390118E+01),
        (lrSetpoint := 2.300000000000000E+02, lrMeasurement := 2.295018207653769E+02, lrOutput := 5.428352658971367E+01, lrITerm := 5.164181552255695E+01),
        (lrSetpoint := 2.300000000000000E+02, lrMeasurement := 2.298579815723359E+02, lrOutput := 4.684615007747561E+01, lrITerm := 5.167732012947297E+01),
        (lrSetpoint := 2.300000000000000E+02, lrMeasurement := 2.297099559641525E+02, lrOutput := 5.524512966148684E+01, lrITerm := 5.174983113843484E+01),
        (lrSetpoint := 2.300000000000000E+02, lrMeasurement := 2.292603224660122E+02, lrOutput := 6.528129601133496E+01, lrITerm := 5.193475052193180E+01),
        (lrSetpoint := 2.300000000000000E+02, lrMeasurement := 2.293897877643200E+02, lrOutput := 5.638338173686626E+01, lrITerm := 5.208730358085180E+01),
        (lrSetpoint := 2.300000000000000E+02, lrMeasurement := 2.292582772953903E+02, lrOutput := 6.019355945087302E+01, lrITerm := 5.227273425700424E+01),
        (lrSetpoint := 2.300000000000000E+02, lrMeasurement := 2.294628253006983E+02, lrOutput := 5.382906615271175E+01, lrITerm := 5.240702793182965E+01),
        (lrSetpoint := 2.300000000000000E+02, lrMeasurement := 2.296473140882134E+02, lrOutput := 5.178979422912075E+01, lrITerm := 5.249519940977629E+01),
        (lrSetpoint := 2.300000000000000E+02, lrMeasurement := 2.298401980923248E+02, lrOutput := 5.002204258732520E+01, lrITerm := 5.253514988669509E+01),
        (lrSetpoint := 2.300000000000000E+02, lrMeasurement := 2.296045205957711E+02, lrOutput := 5.881039040428847E+01, lrITerm := 5.263401973775231E+01),
        (lrSetpoint := 2.300000000000000E+02, lrMeasurement := 2.297323516074078E+02, lrOutput := 5.339932987699066E+01, lrITerm := 5.270093183590035E+01),
        (lrSetpoint := 2.300000000000000E+02, lrMeasurement := 2.296334077365737E+02, lrOutput := 5.701986212258361E+01, lrITerm := 5.279257990175692E+01),
        (lrSetpoint := 2.300000000000000E+02, lrMeasurement := 2.300897704245489E+02, lrOutput := 4.500907971430971E+01, lrITerm := 5.277013729561970E+01),
        (lrSetpoint := 2.300000000000000E+02, lrMeasurement := 2.300498260281075E+02, lrOutput := 5.158960406981092E+01, lrITerm := 5.275768078859282E+01),
        (lrSetpoint := 2.300000000000000E+02, lrMeasurement := 2.302234863296066E+02, lrOutput := 4.798146004656912E+01, lrITerm := 5.270180920619118E+01),
        (lrSetpoint := 2.300000000000000E+02, lrMeasurement := 2.302368370189383E+02, lrOutput := 4.994780106608929E+01, lrITerm := 5.264259995145661E+01),
        (lrSetpoint := 2.300000000000000E+02, lrMeasurement := 2.303656497083887E+02, lrOutput := 4.740496627927007E+01, lrITerm := 5.255118752435943E+01),
        (lrSetpoint := 2.300000000000000E+02, lrMeasurement := 2.300656326678926E+02, lrOutput := 5.636578594658695E+01, lrITerm := 5.253477935738627E+01),
        (lrSetpoint := 2.300000000000000E+02, lrMeasurement := 2.300769671088171E+02, lrOutput := 5.258966324132233E+01, lrITerm := 5.251553758018200E+01),
        (lrSetpoint := 2.300000000000000E+02, lrMeasurement := 2.305703291023916E+02, lrOutput := 4.005450309459560E+01, lrITerm := 5.237295530458411E+01),
        (lrSetpoint := 2.300000000000000E+02, lrMeasurement := 2.299068720312085E+02, lrOutput := 6.220541030787145E+01, lrITerm := 5.239623729678198E+01),
        (lrSetpoint := 2.300000000000000E+02, lrMeasurement := 2.298678125671597E+02, lrOutput := 5.592456489464647E+01, lrITerm := 5.242928415499205E+01),
        (lrSetpoint := 2.300000000000000E+02, lrMeasurement := 2.302592494514098E+02, lrOutput := 4.451504228824698E+01, lrITerm := 5.236447179213961E+01),
        (lrSetpoint := 2.300000000000000E+02, lrMeasurement := 2.303004611033681E+02, lrOutput := 4.807119447949613E+01, lrITerm := 5.228935651629758E+01),
        (lrSetpoint := 2.300000000000000E+02, lrMeasurement := 2.295410621479397E+02, lrOutput := 6.786308244067786E+01, lrITerm := 5.240409097931265E+01),
        (lrSetpoint := 2.300000000000000E+02, lrMeasurement := 2.296394750929767E+02, lrOutput := 5.616131207063897E+01, lrITerm := 5.249422220606846E+01),
        (lrSetpoint := 2.300000000000000E+02, lrMeasurement := 2.297358508945258E+02, lrOutput := 5.328801762312293E+01, lrITerm := 5.256025948243702E+01),
        (lrSetpoint := 2.300000000000000E+02, lrMeasurement := 2.299217984946618E+02, lrOutput := 4.995317335867932E+01, lrITerm := 5.257980985877157E+01),
        (lrSetpoint := 2.300000000000000E+02, lrMeasurement := 2.294578388672089E+02, lrOutput := 6.382554353498379E+01, lrITerm := 5.271535014196933E+01),
        (lrSetpoint := 2.300000000000000E+02, lrMeasurement := 2.295892548900854E+02, lrOutput := 5.535592179887775E+01, lrITerm := 5.281803641944797E+01),
        (lrSetpoint := 2.300000000000000E+02, lrMeasurement := 2.297601347464323E+02, lrOutput := 5.191323195985375E+01, lrITerm := 5.287800273283989E+01),
        (lrSetpoint := 2.300000000000000E+02, lrMeasurement := 2.296982505122999E+02, lrOutput := 5.578084519217992E+01, lrITerm := 5.295344010476492E+01),
        (lrSetpoint := 2.300000000000000E+02, lrMeasurement := 2.295729615193367E+02, lrOutput := 5.856381329480985E+01, lrITerm := 5.306019972493074E+01),
        (lrSetpoint := 2.300000000000000E+02, lrMeasurement := 2.296319668314576E+02, lrOutput := 5.556984951638715E+01, lrITerm := 5.315220801706635E+01),
        (lrSetpoint := 2.300000000000000E+02, lrMeasurement := 2.294668115625297E+02, lrOutput := 6.008817215923838E+01, lrITerm := 5.328550512643393E+01),
        (lrSetpoint := 2.300000000000000E+02, lrMeasurement := 2.296908661859453E+02, lrOutput := 5.275841702434443E+01, lrITerm := 5.336278857994760E+01),
        (lrSetpoint := 2.300000000000000E+02, lrMeasurement := 2.297108953449104E+02, lrOutput := 5.481194702738610E+01, lrITerm := 5.343506474372000E+01),
        (lrSetpoint := 2.300000000000000E+02, lrMeasurement := 2.298020877218476E+02, lrOutput := 5.342157201607348E+01, lrITerm := 5.348454281325811E+01),
        (lrSetpoint := 2.300000000000000E+02, lrMeasurement := 2.296836902792228E+02, lrOutput := 5.765920328718489E+01, lrITerm := 5.356362024345241E+01),
        (lrSetpoint := 2.300000000000000E+02, lrMeasurement := 2.298560098055138E+02, lrOutput := 5.230744798280961E+01, lrITerm := 5.359961779207394E+01),
        (lrSetpoint := 2.300000000000000E+02, lrMeasurement := 2.299300144210812E+02, lrOutput := 5.250410669604547E+01, lrITerm := 5.361711418680364E+01),
        (lrSetpoint := 2.300000000000000E+02, lrMeasurement := 2.297755595039245E+02, lrOutput := 5.760544852951327E+01, lrITerm := 5.367322431082253E+01),
        (lrSetpoint := 2.300000000000000E+02, lrMeasurement := 2.298026433801039E+02, lrOutput := 5.529541445611044E+01, lrITerm := 5.372256346579654E+01),
        (lrSetpoint := 2.300000000000000E+02, lrMeasurement := 2.297567883947042E+02, lrOutput := 5.646153858211288E+01, lrITerm := 5.378336636712050E+01),
        (lrSetpoint := 2.300000000000000E+02, lrMeasurement := 2.297575413877743E+02, lrOutput := 5.591809790338619E+01, lrITerm := 5.384398102017693E+01),
        (lrSetpoint := 2.300000000000000E+02, lrMeasurement := 2.296616659484106E+02, lrOutput := 5.819613357268848E+01, lrITerm := 5.392856453307428E+01),
        (lrSetpoint := 2.300000000000000E+02, lrMeasurement := 2.298497051904085E+02, lrOutput := 5.247204816561817E+01, lrITerm := 5.396613823547216E+01),
        (lrSetpoint := 2.300000000000000E+02, lrMeasurement := 2.297927968721062E+02, lrOutput := 5.604680742411652E+01, lrITerm := 5.401793901744562E+01),
        (lrSetpoint := 2.300000000000000E+02, lrMeasurement := 2.301778769710344E+02, lrOutput := 4.646342110026299E+01, lrITerm := 5.397346977468701E+01),
        (lrSetpoint := 2.300000000000000E+02, lrMeasurement := 2.301251916924390E+02, lrOutput := 5.256619618836143E+01, lrITerm := 5.394217185157725E+01),
        (lrSetpoint := 2.300000000000000E+02, lrMeasurement := 2.299933072438744E+02, lrOutput := 5.603264984190645E+01, lrITerm := 5.394384504060864E+01),
        (lrSetpoint := 2.300000000000000E+02, lrMeasurement := 2.299097613406531E+02, lrOutput := 5.643210098222134E+01, lrITerm := 5.396640470544538E+01),
        (lrSetpoint := 2.300000000000000E+02, lrMeasurement := 2.299827547129346E+02, lrOutput := 5.328954176762921E+01, lrITerm := 5.397071602721172E+01),
        (lrSetpoint := 2.300000000000000E+02, lrMeasurement := 2.304589521651602E+02, lrOutput := 4.240137411780989E+01, lrITerm := 5.385597798592166E+01),
        (lrSetpoint := 2.300000000000000E+02, lrMeasurement := 2.303726599951288E+02, lrOutput := 5.060561043724498E+01, lrITerm := 5.376281298713945E+01),
        (lrSetpoint := 2.300000000000000E+02, lrMeasurement := 2.304580352714455E+02, lrOutput := 4.858283305887362E+01, lrITerm := 5.364830416927807E+01),
        (lrSetpoint := 2.300000000000000E+02, lrMeasurement := 2.301154155085727E+02, lrOutput := 5.789780464175183E+01, lrITerm := 5.361945029213491E+01),
        (lrSetpoint := 2.300000000000000E+02, lrMeasurement := 2.305283091889812E+02, lrOutput := 4.369493628014261E+01, lrITerm := 5.348737299488960E+01),
        (lrSetpoint := 2.300000000000000E+02, lrMeasurement := 2.303795450849513E+02, lrOutput := 5.162315906794111E+01, lrITerm := 5.339248672365179E+01),
        (lrSetpoint := 2.300000000000000E+02, lrMeasurement := 2.300553667625987E+02, lrOutput := 5.837597069463477E+01, lrITerm := 5.337864503300212E+01),
        (lrSetpoint := 2.300000000000000E+02, lrMeasurement := 2.301033416478938E+02, lrOutput := 5.284653022564132E+01, lrITerm := 5.335280962102868E+01),
        (lrSetpoint := 2.300000000000000E+02, lrMeasurement := 2.301573457048873E+02, lrOutput := 5.125473340136315E+01, lrITerm := 5.331347319480685E+01),
        (lrSetpoint := 2.300000000000000E+02, lrMeasurement := 2.300508691127785E+02, lrOutput := 5.443743365725646E+01, lrITerm := 5.330075591661222E+01),
        (lrSetpoint := 2.300000000000000E+02, lrMeasurement := 2.299337282370516E+02, lrOutput := 5.603047810114136E+01, lrITerm := 5.331732385734932E+01),
        (lrSetpoint := 2.300000000000000E+02, lrMeasurement := 2.299160610432337E+02, lrOutput := 5.472909137979824E+01, lrITerm := 5.333830859654088E+01),
        (lrSetpoint := 2.300000000000000E+02, lrMeasurement := 2.298535782085829E+02, lrOutput := 5.568986795597087E+01, lrITerm := 5.337491404439516E+01),
        (lrSetpoint := 2.300000000000000E+02, lrMeasurement := 2.298858958705276E+02, lrOutput := 5.402790643747540E+01, lrITerm := 5.340344007676327E+01),
        (lrSetpoint := 2.300000000000000E+02, lrMeasurement := 2.300523485090222E+02, lrOutput := 5.025064932640316E+01, lrITerm := 5.339035294950772E+01),
        (lrSetpoint := 2.300000000000000E+02, lrMeasurement := 2.293845724968881E+02, lrOutput := 6.860786293414014E+01, lrITerm := 5.354420982528569E+01),
        (lrSetpoint := 2.300000000000000E+02, lrMeasurement := 2.297854823900782E+02, lrOutput := 5.092746843289019E+01, lrITerm := 5.359783922776613E+01),
        (lrSetpoint := 2.300000000000000E+02, lrMeasurement := 2.298561685559700E+02, lrOutput := 5.277616765189516E+01, lrITerm := 5.363379708877363E+01),
        (lrSetpoint := 2.300000000000000E+02, lrMeasurement := 2.298627366738675E+02, lrOutput := 5.425947344518362E+01, lrITerm := 5.366811292030675E+01),
        (lrSetpoint := 2.300000000000000E+02, lrMeasurement := 2.297464639181015E+02, lrOutput := 5.751880047138757E+01, lrITerm := 5.373149694078137E+01),
        (lrSetpoint := 2.300000000000000E+02, lrMeasurement := 2.295433810930751E+02, lrOutput := 6.109973109841962E+01, lrITerm := 5.384565166751261E+01),
        (lrSetpoint := 2.300000000000000E+02, lrMeasurement := 2.299039995658953E+02, lrOutput := 4.958798531885385E+01, lrITerm := 5.386965177603878E+01)
    ];
    aWestgard : ARRAY[1..300] OF ST_WestgardVector := [
        (diStep := 0, lrValue := 2.504570756196317E+01, bWarn12s := FALSE, bReject13s := FALSE, bReject22s := FALSE),
        (diStep := 1, lrValue := 2.559400238406393E+01, bWarn12s := FALSE, bReject13s := FALSE, bReject22s := FALSE),
        (diStep := 2, lrValue := 2.721106767937097E+01, bWarn12s := FALSE, bReject13s := FALSE, bReject22s := FALSE),
        (diStep := 3, lrValue := 2.906538770745868E+01, bWarn12s := FALSE, bReject13s := FALSE, bReject22s := FALSE),
        (diStep := 4, lrValue := 3.083779911570193E+01, bWarn12s := FALSE, bReject13s := FALSE, bReject22s := FALSE),
        (diStep := 5, lrValue := 3.344406655918265E+01, bWarn12s := FALSE, bReject13s := FALSE, bReject22s := FALSE),
        (diStep := 6, lrValue := 3.640825075871666E+01, bWarn12s := FALSE, bReject13s := FALSE, bReject22s := FALSE),
        (diStep := 7, lrValue := 3.928242815999355E+01, bWarn12s := FALSE, bReject13s := FALSE, bReject22s := FALSE),
        (diStep := 8, lrValue := 4.241953904612176E+01, bWarn12s := FALSE, bReject13s := FALSE, bReject22s := FALSE),
        (diStep := 9, lrValue := 4.550594203217187E+01, bWarn12s := FALSE, bReject13s := FALSE, bReject22s := FALSE),
        (diStep := 10, lrValue := 4.907188733629471E+01, bWarn12s := FALSE, bReject13s := FALSE, bReject22s := FALSE),
        (diStep := 11, lrValue := 5.243664392789950E+01, bWarn12s := FALSE, bReject13s := FALSE, bReject22s := FALSE),
        (diStep := 12, lrValue := 5.576754175418417E+01, bWarn12s := FALSE, bReject13s := FALSE, bReject22s := FALSE),
        (diStep := 13, lrValue := 5.940904962608809E+01, bWarn12s := FALSE, bReject13s := FALSE, bReject22s := FALSE),
        (diStep := 14, lrValue := 6.282668317532421E+01, bWarn12s := FALSE, bReject13s := FALSE, bReject22s := FALSE),
        (diStep := 15, lrValue := 6.617020839567282E+01, bWarn12s := FALSE, bReject13s := FALSE, bReject22s := FALSE),
        (diStep := 16, lrValue := 6.991626356192097E+01, bWarn12s := FALSE, bReject13s := FALSE, bReject22s := FALSE),
        (diStep := 17, lrValue := 7.329295415928244E+01, bWarn12s := FALSE, bReject13s := FALSE, bReject22s := FALSE),
        (diStep := 18, lrValue := 7.715412652709350E+01, bWarn12s := FALSE, bReject13s := FALSE, bReject22s := FALSE),
        (diStep := 19, lrValue := 8.060678218175724E+01, bWarn12s := FALSE, bReject13s := FALSE, bReject22s := FALSE),
        (diStep := 20, lrValue := 8.418207861531381E+01, bWarn12s := FALSE, bReject13s := FALSE, bReject22s := FALSE),
        (diStep := 21, lrValue := 8.770466127710711E+01, bWarn12s := FALSE, bReject13s := FALSE, bReject22s := FALSE),
        (diStep := 22, lrValue := 9.158689819204071E+01, bWarn12s := FALSE, bReject13s := FALSE, bReject22s := FALSE),
        (diStep := 23, lrValue := 9.497539444205835E+01, bWarn12s := FALSE, bReject13s := FALSE, bReject22s := FALSE),
        (diStep := 24, lrValue := 9.852661866900469E+01, bWarn12s := FALSE, bReject13s := FALSE, bReject22s := FALSE),
        (diStep := 25, lrValue := 1.021266989746227E+02, bWarn12s := FALSE, bReject13s := FALSE, bReject22s := FALSE),
        (diStep := 26, lrValue := 1.058436726674556E+02, bWarn12s := FALSE, bReject13s := FALSE, bReject22s := FALSE),
        (diStep := 27, lrValue := 1.093980483030509E+02, bWarn12s := FALSE, bReject13s := FALSE, bReject22s := FALSE),
        (diStep := 28, lrValue := 1.129792015668312E+02, bWarn12s := FALSE, bReject13s := FALSE, bReject22s := FALSE),
        (diStep := 29, lrValue := 1.165502773982586E+02, bWarn12s := FALSE, bReject13s := FALSE, bReject22s := FALSE),
        (diStep := 30, lrValue := 1.203692878042951E+02, bWarn12s := FALSE, bReject13s := FALSE, bReject22s := FALSE),
        (diStep := 31, lrValue := 1.235432685102606E+02, bWarn12s := FALSE, bReject13s := FALSE, bReject22s := FALSE),
        (diStep := 32, lrValue := 1.270772148357379E+02, bWarn12s := FALSE, bReject13s := FALSE, bReject22s := FALSE),
        (diStep := 33, lrValue := 1.305753003884958E+02, bWarn12s := FALSE, bReject13s := FALSE, bReject22s := FALSE),
        (diStep := 34, lrValue := 1.343264670026235E+02, bWarn12s := FALSE, bReject13s := FALSE, bReject22s := FALSE),
        (diStep := 35, lrValue := 1.379334266122466E+02, bWarn12s := FALSE, bReject13s := FALSE, bReject22s := FALSE),
        (diStep := 36, lrValue := 1.412702435435773E+02, bWarn12s := FALSE, bReject13s := FALSE, bReject22s := FALSE),
        (diStep := 37, lrValue := 1.446777639636957E+02, bWarn12s := FALSE, bReject13s := FALSE, bReject22s := FALSE),
        (diStep := 38, lrValue := 1.481897288334872E+02, bWarn12s := FALSE, bReject13s := FALSE, bReject22s := FALSE),
        (diStep := 39, lrValue := 1.519137400563598E+02, bWarn12s := FALSE, bReject13s := FALSE, bReject22s := FALSE),
        (diStep := 40, lrValue := 1.554235085010919E+02, bWarn12s := FALSE, bReject13s := FALSE, bReject22s := FALSE),
        (diStep := 41, lrValue := 1.588824707065076E+02, bWarn12s := FALSE, bReject13s := FALSE, bReject22s := FALSE),
        (diStep := 42, lrValue := 1.621832501003170E+02, bWarn12s := FALSE, bReject13s := FALSE, bReject22s := FALSE),
        (diStep := 43, lrValue := 1.657930793899823E+02, bWarn12s := FALSE, bReject13s := FALSE, bReject22s := FALSE),
        (diStep := 44, lrValue := 1.692440373830902E+02, bWarn12s := FALSE, bReject13s := FALSE, bReject22s := FALSE),
        (diStep := 45, lrValue := 1.727207213966689E+02, bWarn12s := FALSE, bReject13s := FALSE, bReject22s := FALSE),
        (diStep := 46, lrValue := 1.762731259192086E+02, bWarn12s := FALSE, bReject13s := FALSE, bReject22s := FALSE),
        (diStep := 47, lrValue := 1.796235615768844E+02, bWarn12s := FALSE, bReject13s := FALSE, bReject22s := FALSE),
        (diStep := 48, lrValue := 1.831325956067453E+02, bWarn12s := FALSE, bReject13s := FALSE, bReject22s := FALSE),
        (diStep := 49, lrValue := 1.864747670133277E+02, bWarn12s := FALSE, bReject13s := FALSE, bReject22s := FALSE),
        (diStep := 50, lrValue := 1.899350152806136E+02, bWarn12s := FALSE, bReject13s := FALSE, bReject22s := FALSE),
        (diStep := 51, lrValue := 1.934065144925135E+02, bWarn12s := FALSE, bReject13s := FALSE, bReject22s := FALSE),
        (diStep := 52, lrValue := 1.965065899891975E+02, bWarn12s := FALSE, bReject13s := FALSE, bReject22s := FALSE),
        (diStep := 53, lrValue := 2.000837349498422E+02, bWarn12s := FALSE, bReject13s := FALSE, bReject22s := FALSE),
        (diStep := 54, lrValue := 2.034608444403627E+02, bWarn12s := FALSE, bReject13s := FALSE, bReject22s := FALSE),
        (diStep := 55, lrValue := 2.068284883225735E+02, bWarn12s := FALSE, bReject13s := FALSE, bReject22s := FALSE),
        (diStep := 56, lrValue := 2.102691859917106E+02, bWarn12s := FALSE, bReject13s := FALSE, bReject22s := FALSE),
        (diStep := 57, lrValue := 2.138707975791627E+02, bWarn12s := FALSE, bReject13s := FALSE, bReject22s := FALSE),
        (diStep := 58, lrValue := 2.166047382771748E+02, bWarn12s := FALSE, bReject13s := FALSE, bReject22s := FALSE),
        (diStep := 59, lrValue := 2.196531259180408E+02, bWarn12s := FALSE, bReject13s := FALSE, bReject22s := FALSE),
        (diStep := 60, lrValue := 2.215944746720401E+02, bWarn12s := FALSE, bReject13s := FALSE, bReject22s := FALSE),
        (diStep := 61, lrValue := 2.238164015632227E+02, bWarn12s := FALSE, bReject13s := FALSE, bReject22s := FALSE),
        (diStep := 62, lrValue := 2.255252359017419E+02, bWarn12s := FALSE, bReject13s := FALSE, bReject22s := FALSE),
        (diStep := 63, lrValue := 2.268803103257552E+02, bWarn12s := FALSE, bReject13s := FALSE, bReject22s := FALSE),
        (diStep := 64, lrValue := 2.278955664907341E+02, bWarn12s := FALSE, bReject13s := FALSE, bReject22s := FALSE),
        (diStep := 65, lrValue := 2.286631929043172E+02, bWarn12s := FALSE, bReject13s := FALSE, bReject22s := FALSE),
        (diStep := 66, lrValue := 2.290508932078158E+02, bWarn12s := FALSE, bReject13s := FALSE, bReject22s := FALSE),
        (diStep := 67, lrValue := 2.294681164603311E+02, bWarn12s := FALSE, bReject13s := FALSE, bReject22s := FALSE),
        (diStep := 68, lrValue := 2.299838292420773E+02, bWarn12s := FALSE, bReject13s := FALSE, bReject22s := FALSE),
        (diStep := 69, lrValue := 2.300096375187556E+02, bWarn12s := FALSE, bReject13s := FALSE, bReject22s := FALSE),
        (diStep := 70, lrValue := 2.299780300469962E+02, bWarn12s := FALSE, bReject13s := FALSE, bReject22s := FALSE),
        (diStep := 71, lrValue := 2.301089493703319E+02, bWarn12s := FALSE, bReject13s := FALSE, bReject22s := FALSE),
        (diStep := 72, lrValue := 2.302094572798513E+02, bWarn12s := FALSE, bReject13s := FALSE, bReject22s := FALSE),
        (diStep := 73, lrValue := 2.304978744922259E+02, bWarn12s := FALSE, bReject13s := FALSE, bReject22s := FALSE),
        (diStep := 74, lrValue := 2.304858332660471E+02, bWarn12s := FALSE, bReject13s := FALSE, bReject22s := FALSE),
        (diStep := 75, lrValue := 2.306128359144820E+02, bWarn12s := FALSE, bReject13s := FALSE, bReject22s := FALSE),
        (diStep := 76, lrValue := 2.304736944247048E+02, bWarn12s := FALSE, bReject13s := FALSE, bReject22s := FALSE),
        (diStep := 77, lrValue := 2.306144061359000E+02, bWarn12s := FALSE, bReject13s := FALSE, bReject22s := FALSE),
        (diStep := 78, lrValue := 2.307194784114588E+02, bWarn12s := FALSE, bReject13s := FALSE, bReject22s := FALSE),
        (diStep := 79, lrValue := 2.305911113626528E+02, bWarn12s := FALSE, bReject13s := FALSE, bReject22s := FALSE),
        (diStep := 80, lrValue := 2.307337919192282E+02, bWarn12s := FALSE, bReject13s := FALSE, bReject22s := FALSE),
        (diStep := 81, lrValue := 2.305232005023320E+02, bWarn12s := FALSE, bReject13s := FALSE, bReject22s := FALSE),
        (diStep := 82, lrValue := 2.305177106373760E+02, bWarn12s := FALSE, bReject13s := FALSE, bReject22s := FALSE),
        (diStep := 83, lrValue := 2.304407682616513E+02, bWarn12s := FALSE, bReject13s := FALSE, bReject22s := FALSE),
        (diStep := 84, lrValue := 2.302345111439646E+02, bWarn12s := FALSE, bReject13s := FALSE, bReject22s := FALSE),
        (diStep := 85, lrValue := 2.304233655001475E+02, bWarn12s := FALSE, bReject13s := FALSE, bReject22s := FALSE),
        (diStep := 86, lrValue := 2.301765571888204E+02, bWarn12s := FALSE, bReject13s := FALSE, bReject22s := FALSE),
        (diStep := 87, lrValue := 2.301718013630896E+02, bWarn12s := FALSE, bReject13s := FALSE, bReject22s := FALSE),
        (diStep := 88, lrValue := 2.301656351697725E+02, bWarn12s := FALSE, bReject13s := FALSE, bReject22s := FALSE),
        (diStep := 89, lrValue := 2.300808227245562E+02, bWarn12s := FALSE, bReject13s := FALSE, bReject22s := FALSE),
        (diStep := 90, lrValue := 2.300450161809068E+02, bWarn12s := FALSE, bReject13s := FALSE, bReject22s := FALSE),
        (diStep := 91, lrValue := 2.298685710227648E+02, bWarn12s := FALSE, bReject13s := FALSE, bReject22s := FALSE),
        (diStep := 92, lrValue := 2.297903074584952E+02, bWarn12s := FALSE, bReject13s := FALSE, bReject22s := FALSE),
        (diStep := 93, lrValue := 2.298346004226570E+02, bWarn12s := FALSE, bReject13s := FALSE, bReject22s := FALSE),
        (diStep := 94, lrValue := 2.295852197770309E+02, bWarn12s := FALSE, bReject13s := FALSE, bReject22s := FALSE),
        (diStep := 95, lrValue := 2.296599261274224E+02, bWarn12s := FALSE, bReject13s := FALSE, bReject22s := FALSE),
        (diStep := 96, lrValue := 2.297182708644902E+02, bWarn12s := FALSE, bReject13s := FALSE, bReject22s := FALSE),
        (diStep := 97, lrValue := 2.298000366341335E+02, bWarn12s := FALSE, bReject13s := FALSE, bReject22s := FALSE),
        (diStep := 98, lrValue := 2.300288961980845E+02, bWarn12s := FALSE, bReject13s := FALSE, bReject22s := FALSE),
        (diStep := 99, lrValue := 2.298093482091375E+02, bWarn12s := FALSE, bReject13s := FALSE, bReject22s := FALSE),
        (diStep := 100, lrValue := 2.298940447799201E+02, bWarn12s := FALSE, bReject13s := FALSE, bReject22s := FALSE),
        (diStep := 101, lrValue := 2.301432779377677E+02, bWarn12s := FALSE, bReject13s := FALSE, bReject22s := FALSE),
        (diStep := 102, lrValue := 2.298459618394776E+02, bWarn12s := FALSE, bReject13s := FALSE, bReject22s := FALSE),
        (diStep := 103, lrValue := 2.300026310488091E+02, bWarn12s := FALSE, bReject13s := FALSE, bReject22s := FALSE),
        (diStep := 104, lrValue := 2.297259479761731E+02, bWarn12s := FALSE, bReject13s := FALSE, bReject22s := FALSE),
        (diStep := 105, lrValue := 2.298549920521735E+02, bWarn12s := FALSE, bReject13s := FALSE, bReject22s := FALSE),
        (diStep := 106, lrValue := 2.297521760524508E+02, bWarn12s := FALSE, bReject13s := FALSE, bReject22s := FALSE),
        (diStep := 107, lrValue := 2.298704273997785E+02, bWarn12s := FALSE, bReject13s := FALSE, bReject22s := FALSE),
        (diStep := 108, lrValue := 2.300586262338561E+02, bWarn12s := FALSE, bReject13s := FALSE, bReject22s := FALSE),
        (diStep := 109, lrValue := 2.296482659229140E+02, bWarn12s := FALSE, bReject13s := FALSE, bReject22s := FALSE),
        (diStep := 110, lrValue := 2.300127602678513E+02, bWarn12s := FALSE, bReject13s := FALSE, bReject22s := FALSE),
        (diStep := 111, lrValue := 2.299745877595838E+02, bWarn12s := FALSE, bReject13s := FALSE, bReject22s := FALSE),
        (diStep := 112, lrValue := 2.298370036522997E+02, bWarn12s := FALSE, bReject13s := FALSE, bReject22s := FALSE),
        (diStep := 113, lrValue := 2.297662189294558E+02, bWarn12s := FALSE, bReject13s := FALSE, bReject22s := FALSE),
        (diStep := 114, lrValue := 2.301069608762478E+02, bWarn12s := FALSE, bReject13s := FALSE, bReject22s := FALSE),
        (diStep := 115, lrValue := 2.301034615741697E+02, bWarn12s := FALSE, bReject13s := FALSE, bReject22s := FALSE),
        (diStep := 116, lrValue := 2.303148002423178E+02, bWarn12s := FALSE, bReject13s := FALSE, bReject22s := FALSE),
        (diStep := 117, lrValue := 2.303555301449315E+02, bWarn12s := FALSE, bReject13s := FALSE, bReject22s := FALSE),
        (diStep := 118, lrValue := 2.306586161636685E+02, bWarn12s := FALSE, bReject13s := FALSE, bReject22s := FALSE),
        (diStep := 119, lrValue := 2.303959258597061E+02, bWarn12s := FALSE, bReject13s := FALSE, bReject22s := FALSE),
        (diStep := 120, lrValue := 2.303270774525105E+02, bWarn12s := FALSE, bReject13s := FALSE, bReject22s := FALSE),
        (diStep := 121, lrValue := 2.305308276598897E+02, bWarn12s := FALSE, bReject13s := FALSE, bReject22s := FALSE),
        (diStep := 122, lrValue := 2.304918859423371E+02, bWarn12s := FALSE, bReject13s := FALSE, bReject22s := FALSE),
        (diStep := 123, lrValue := 2.305868168294902E+02, bWarn12s := TRUE, bReject13s := FALSE, bReject22s := FALSE),
        (diStep := 124, lrValue := 2.303892627913187E+02, bWarn12s := FALSE, bReject13s := FALSE, bReject22s := FALSE),
        (diStep := 125, lrValue := 2.302083083202458E+02, bWarn12s := FALSE, bReject13s := FALSE, bReject22s := FALSE),
        (diStep := 126, lrValue := 2.302879174462091E+02, bWarn12s := FALSE, bReject13s := FALSE, bReject22s := FALSE),
        (diStep := 127, lrValue := 2.297863666250582E+02, bWarn12s := FALSE, bReject13s := FALSE, bReject22s := FALSE),
        (diStep := 128, lrValue := 2.298453652638796E+02, bWarn12s := FALSE, bReject13s := FALSE, bReject22s := FALSE),
        (diStep := 129, lrValue := 2.297852853998048E+02, bWarn12s := FALSE, bReject13s := FALSE, bReject22s := FALSE),
        (diStep := 130, lrValue := 2.298611656666668E+02, bWarn12s := FALSE, bReject13s := FALSE, bReject22s := FALSE),
        (diStep := 131, lrValue := 2.296984707598905E+02, bWarn12s := FALSE, bReject13s := FALSE, bReject22s := FALSE),
        (diStep := 132, lrValue := 2.300134306392112E+02, bWarn12s := FALSE, bReject13s := FALSE, bReject22s := FALSE),
        (diStep := 133, lrValue := 2.298490494877590E+02, bWarn12s := FALSE, bReject13s := FALSE, bReject22s := FALSE),
        (diStep := 134, lrValue := 2.296442219691345E+02, bWarn12s := FALSE, bReject13s := FALSE, bReject22s := FALSE),
        (diStep := 135, lrValue := 2.297367369885094E+02, bWarn12s := FALSE, bReject13s := FALSE, bReject22s := FALSE),
        (diStep := 136, lrValue := 2.299557157451501E+02, bWarn12s := FALSE, bReject13s := FALSE, bReject22s := FALSE),
        (diStep := 137, lrValue := 2.300155318818599E+02, bWarn12s := FALSE, bReject13s := FALSE, bReject22s := FALSE),
        (diStep := 138, lrValue := 2.301509214398248E+02, bWarn12s := FALSE, bReject13s := FALSE, bReject22s := FALSE),
        (diStep := 139, lrValue := 2.302200352161047E+02, bWarn12s := FALSE, bReject13s := FALSE, bReject22s := FALSE),
        (diStep := 140, lrValue := 2.297549336201718E+02, bWarn12s := FALSE, bReject13s := FALSE, bReject22s := FALSE),
        (diStep := 141, lrValue := 2.295307302659245E+02, bWarn12s := FALSE, bReject13s := FALSE, bReject22s := FALSE),
        (diStep := 142, lrValue := 2.294052885678543E+02, bWarn12s := TRUE, bReject13s := FALSE, bReject22s := FALSE),
        (diStep := 143, lrValue := 2.298522298602363E+02, bWarn12s := FALSE, bReject13s := FALSE, bReject22s := FALSE),
        (diStep := 144, lrValue := 2.297115211052058E+02, bWarn12s := FALSE, bReject13s := FALSE, bReject22s := FALSE),
        (diStep := 145, lrValue := 2.298054273966737E+02, bWarn12s := FALSE, bReject13s := FALSE, bReject22s := FALSE),
        (diStep := 146, lrValue := 2.297982350513737E+02, bWarn12s := FALSE, bReject13s := FALSE, bReject22s := FALSE),
        (diStep := 147, lrValue := 2.298912673017996E+02, bWarn12s := FALSE, bReject13s := FALSE, bReject22s := FALSE),
        (diStep := 148, lrValue := 2.300789608336171E+02, bWarn12s := FALSE, bReject13s := FALSE, bReject22s := FALSE),
        (diStep := 149, lrValue := 2.299119910387465E+02, bWarn12s := FALSE, bReject13s := FALSE, bReject22s := FALSE),
        (diStep := 150, lrValue := 2.298543613889811E+02, bWarn12s := FALSE, bReject13s := FALSE, bReject22s := FALSE),
        (diStep := 151, lrValue := 2.294720232167521E+02, bWarn12s := FALSE, bReject13s := FALSE, bReject22s := FALSE),
        (diStep := 152, lrValue := 2.289971171519480E+02, bWarn12s := FALSE, bReject13s := TRUE, bReject22s := FALSE),
        (diStep := 153, lrValue := 2.287900661865506E+02, bWarn12s := FALSE, bReject13s := TRUE, bReject22s := TRUE),
        (diStep := 154, lrValue := 2.284515985235186E+02, bWarn12s := FALSE, bReject13s := TRUE, bReject22s := TRUE),
        (diStep := 155, lrValue := 2.283411627174421E+02, bWarn12s := FALSE, bReject13s := TRUE, bReject22s := TRUE),
        (diStep := 156, lrValue := 2.277124386479682E+02, bWarn12s := FALSE, bReject13s := TRUE, bReject22s := TRUE),
        (diStep := 157, lrValue := 2.275574921917000E+02, bWarn12s := FALSE, bReject13s := TRUE, bReject22s := TRUE),
        (diStep := 158, lrValue := 2.271008315546960E+02, bWarn12s := FALSE, bReject13s := TRUE, bReject22s := TRUE),
        (diStep := 159, lrValue := 2.268624201050854E+02, bWarn12s := FALSE, bReject13s := TRUE, bReject22s := TRUE),
        (diStep := 160, lrValue := 2.268378562653796E+02, bWarn12s := FALSE, bReject13s := TRUE, bReject22s := TRUE),
        (diStep := 161, lrValue := 2.268104966628377E+02, bWarn12s := FALSE, bReject13s := TRUE, bReject22s := TRUE),
        (diStep := 162, lrValue := 2.271727202882387E+02, bWarn12s := FALSE, bReject13s := TRUE, bReject22s := TRUE),
        (diStep := 163, lrValue := 2.265982553891899E+02, bWarn12s := FALSE, bReject13s := TRUE, bReject22s := TRUE),
        (diStep := 164, lrValue := 2.268067431131597E+02, bWarn12s := FALSE, bReject13s := TRUE, bReject22s := TRUE),
        (diStep := 165, lrValue := 2.264977102339018E+02, bWarn12s := FALSE, bReject13s := TRUE, bReject22s := TRUE),
        (diStep := 166, lrValue := 2.267918815203126E+02, bWarn12s := FALSE, bReject13s := TRUE, bReject22s := TRUE),
        (diStep := 167, lrValue := 2.267072664589627E+02, bWarn12s := FALSE, bReject13s := TRUE, bReject22s := TRUE),
        (diStep := 168, lrValue := 2.266504042455074E+02, bWarn12s := FALSE, bReject13s := TRUE, bReject22s := TRUE),
        (diStep := 169, lrValue := 2.267264485475885E+02, bWarn12s := FALSE, bReject13s := TRUE, bReject22s := TRUE),
        (diStep := 170, lrValue := 2.267063455066636E+02, bWarn12s := FALSE, bReject13s := TRUE, bReject22s := TRUE),
        (diStep := 171, lrValue := 2.269697698730993E+02, bWarn12s := FALSE, bReject13s := TRUE, bReject22s := TRUE),
        (diStep := 172, lrValue := 2.269111095789345E+02, bWarn12s := FALSE, bReject13s := TRUE, bReject22s := TRUE),
        (diStep := 173, lrValue := 2.268960923785198E+02, bWarn12s := FALSE, bReject13s := TRUE, bReject22s := TRUE),
        (diStep := 174, lrValue := 2.270156326598504E+02, bWarn12s := FALSE, bReject13s := TRUE, bReject22s := TRUE),
        (diStep := 175, lrValue := 2.273641290287552E+02, bWarn12s := FALSE, bReject13s := TRUE, bReject22s := TRUE),
        (diStep := 176, lrValue := 2.276619484977107E+02, bWarn12s := FALSE, bReject13s := TRUE, bReject22s := TRUE),
        (diStep := 177, lrValue := 2.274873010596821E+02, bWarn12s := FALSE, bReject13s := TRUE, bReject22s := TRUE),
        (diStep := 178, lrValue := 2.275169921363721E+02, bWarn12s := FALSE, bReject13s := TRUE, bReject22s := TRUE),
        (diStep := 179, lrValue := 2.276650690346880E+02, bWarn12s := FALSE, bReject13s := TRUE, bReject22s := TRUE),
        (diStep := 180, lrValue := 2.278966070310045E+02, bWarn12s := FALSE, bReject13s := TRUE, bReject22s := TRUE),
        (diStep := 181, lrValue := 2.277815965043510E+02, bWarn12s := FALSE, bReject13s := TRUE, bReject22s := TRUE),
        (diStep := 182, lrValue := 2.277607171447250E+02, bWarn12s := FALSE, bReject13s := TRUE, bReject22s := TRUE),
        (diStep := 183, lrValue := 2.280841211516531E+02, bWarn12s := FALSE, bReject13s := TRUE, bReject22s := TRUE),
        (diStep := 184, lrValue := 2.280378619566982E+02, bWarn12s := FALSE, bReject13s := TRUE, bReject22s := TRUE),
        (diStep := 185, lrValue := 2.282695321084727E+02, bWarn12s := FALSE, bReject13s := TRUE, bReject22s := TRUE),
        (diStep := 186, lrValue := 2.281034579844685E+02, bWarn12s := FALSE, bReject13s := TRUE, bReject22s := TRUE),
        (diStep := 187, lrValue := 2.279622185203662E+02, bWarn12s := FALSE, bReject13s := TRUE, bReject22s := TRUE),
        (diStep := 188, lrValue := 2.280545056773856E+02, bWarn12s := FALSE, bReject13s := TRUE, bReject22s := TRUE),
        (diStep := 189, lrValue := 2.286269974803834E+02, bWarn12s := FALSE, bReject13s := TRUE, bReject22s := TRUE),
        (diStep := 190, lrValue := 2.286671160554017E+02, bWarn12s := FALSE, bReject13s := TRUE, bReject22s := TRUE),
        (diStep := 191, lrValue := 2.283905080974753E+02, bWarn12s := FALSE, bReject13s := TRUE, bReject22s := TRUE),
        (diStep := 192, lrValue := 2.284205711481603E+02, bWarn12s := FALSE, bReject13s := TRUE, bReject22s := TRUE),
        (diStep := 193, lrValue := 2.288186192176935E+02, bWarn12s := FALSE, bReject13s := TRUE, bReject22s := TRUE),
        (diStep := 194, lrValue := 2.285314344307211E+02, bWarn12s := FALSE, bReject13s := TRUE, bReject22s := TRUE),
        (diStep := 195, lrValue := 2.287350459843640E+02, bWarn12s := FALSE, bReject13s := TRUE, bReject22s := TRUE),
        (diStep := 196, lrValue := 2.291414097941779E+02, bWarn12s := TRUE, bReject13s := FALSE, bReject22s := TRUE),
        (diStep := 197, lrValue := 2.291081848729324E+02, bWarn12s := FALSE, bReject13s := TRUE, bReject22s := TRUE),
        (diStep := 198, lrValue := 2.292964414262748E+02, bWarn12s := TRUE, bReject13s := FALSE, bReject22s := TRUE),
        (diStep := 199, lrValue := 2.293808272853664E+02, bWarn12s := TRUE, bReject13s := FALSE, bReject22s := TRUE),
        (diStep := 200, lrValue := 2.295518096900797E+02, bWarn12s := FALSE, bReject13s := FALSE, bReject22s := FALSE),
        (diStep := 201, lrValue := 2.297340947421611E+02, bWarn12s := FALSE, bReject13s := FALSE, bReject22s := FALSE),
        (diStep := 202, lrValue := 2.294861354096551E+02, bWarn12s := FALSE, bReject13s := FALSE, bReject22s := FALSE),
        (diStep := 203, lrValue := 2.295284263331895E+02, bWarn12s := FALSE, bReject13s := FALSE, bReject22s := FALSE),
        (diStep := 204, lrValue := 2.290650907176098E+02, bWarn12s := FALSE, bReject13s := TRUE, bReject22s := FALSE),
        (diStep := 205, lrValue := 2.293768370143731E+02, bWarn12s := TRUE, bReject13s := FALSE, bReject22s := TRUE),
        (diStep := 206, lrValue := 2.292258378088339E+02, bWarn12s := TRUE, bReject13s := FALSE, bReject22s := TRUE),
        (diStep := 207, lrValue := 2.291530512192492E+02, bWarn12s := TRUE, bReject13s := FALSE, bReject22s := TRUE),
        (diStep := 208, lrValue := 2.292043165056924E+02, bWarn12s := TRUE, bReject13s := FALSE, bReject22s := TRUE),
        (diStep := 209, lrValue := 2.292824733439275E+02, bWarn12s := TRUE, bReject13s := FALSE, bReject22s := TRUE),
        (diStep := 210, lrValue := 2.294540619211454E+02, bWarn12s := FALSE, bReject13s := FALSE, bReject22s := FALSE),
        (diStep := 211, lrValue := 2.290702146383318E+02, bWarn12s := FALSE, bReject13s := TRUE, bReject22s := FALSE),
        (diStep := 212, lrValue := 2.292902545832142E+02, bWarn12s := TRUE, bReject13s := FALSE, bReject22s := TRUE),
        (diStep := 213, lrValue := 2.292086951375199E+02, bWarn12s := TRUE, bReject13s := FALSE, bReject22s := TRUE),
        (diStep := 214, lrValue := 2.292419763819967E+02, bWarn12s := TRUE, bReject13s := FALSE, bReject22s := TRUE),
        (diStep := 215, lrValue := 2.294530367481974E+02, bWarn12s := FALSE, bReject13s := FALSE, bReject22s := FALSE),
        (diStep := 216, lrValue := 2.293613959075460E+02, bWarn12s := TRUE, bReject13s := FALSE, bReject22s := FALSE),
        (diStep := 217, lrValue := 2.294712797684037E+02, bWarn12s := FALSE, bReject13s := FALSE, bReject22s := FALSE),
        (diStep := 218, lrValue := 2.292235190820188E+02, bWarn12s := TRUE, bReject13s := FALSE, bReject22s := FALSE),
        (diStep := 219, lrValue := 2.291629751724858E+02, bWarn12s := TRUE, bReject13s := FALSE, bReject22s := TRUE),
        (diStep := 220, lrValue := 2.292804089571940E+02, bWarn12s := TRUE, bReject13s := FALSE, bReject22s := TRUE),
        (diStep := 221, lrValue := 2.293874877761780E+02, bWarn12s := TRUE, bReject13s := FALSE, bReject22s := TRUE),
        (diStep := 222, lrValue := 2.293982407687014E+02, bWarn12s := TRUE, bReject13s := FALSE, bReject22s := TRUE),
        (diStep := 223, lrValue := 2.292279554865906E+02, bWarn12s := TRUE, bReject13s := FALSE, bReject22s := TRUE),
        (diStep := 224, lrValue := 2.294571546504262E+02, bWarn12s := FALSE, bReject13s := FALSE, bReject22s := FALSE),
        (diStep := 225, lrValue := 2.295018207653769E+02, bWarn12s := FALSE, bReject13s := FALSE, bReject22s := FALSE),
        (diStep := 226, lrValue := 2.298579815723359E+02, bWarn12s := FALSE, bReject13s := FALSE, bReject22s := FALSE),
        (diStep := 227, lrValue := 2.297099559641525E+02, bWarn12s := FALSE, bReject13s := FALSE, bReject22s := FALSE),
        (diStep := 228, lrValue := 2.292603224660122E+02, bWarn12s := TRUE, bReject13s := FALSE, bReject22s := FALSE),
        (diStep := 229, lrValue := 2.293897877643200E+02, bWarn12s := TRUE, bReject13s := FALSE, bReject22s := TRUE),
        (diStep := 230, lrValue := 2.292582772953903E+02, bWarn12s := TRUE, bReject13s := FALSE, bReject22s := TRUE),
        (diStep := 231, lrValue := 2.294628253006983E+02, bWarn12s := FALSE, bReject13s := FALSE, bReject22s := FALSE),
        (diStep := 232, lrValue := 2.296473140882134E+02, bWarn12s := FALSE, bReject13s := FALSE, bReject22s := FALSE),
        (diStep := 233, lrValue := 2.298401980923248E+02, bWarn12s := FALSE, bReject13s := FALSE, bReject22s := FALSE),
        (diStep := 234, lrValue := 2.296045205957711E+02, bWarn12s := FALSE, bReject13s := FALSE, bReject22s := FALSE),
        (diStep := 235, lrValue := 2.297323516074078E+02, bWarn12s := FALSE, bReject13s := FALSE, bReject22s := FALSE),
        (diStep := 236, lrValue := 2.296334077365737E+02, bWarn12s := FALSE, bReject13s := FALSE, bReject22s := FALSE),
        (diStep := 237, lrValue := 2.300897704245489E+02, bWarn12s := FALSE, bReject13s := FALSE, bReject22s := FALSE),
        (diStep := 238, lrValue := 2.300498260281075E+02, bWarn12s := FALSE, bReject13s := FALSE, bReject22s := FALSE),
        (diStep := 239, lrValue := 2.302234863296066E+02, bWarn12s := FALSE, bReject13s := FALSE, bReject22s := FALSE),
        (diStep := 240, lrValue := 2.302368370189383E+02, bWarn12s := FALSE, bReject13s := FALSE, bReject22s := FALSE),
        (diStep := 241, lrValue := 2.303656497083887E+02, bWarn12s := FALSE, bReject13s := FALSE, bReject22s := FALSE),
        (diStep := 242, lrValue := 2.300656326678926E+02, bWarn12s := FALSE, bReject13s := FALSE, bReject22s := FALSE),
        (diStep := 243, lrValue := 2.300769671088171E+02, bWarn12s := FALSE, bReject13s := FALSE, bReject22s := FALSE),
        (diStep := 244, lrValue := 2.305703291023916E+02, bWarn12s := FALSE, bReject13s := FALSE, bReject22s := FALSE),
        (diStep := 245, lrValue := 2.299068720312085E+02, bWarn12s := FALSE, bReject13s := FALSE, bReject22s := FALSE),
        (diStep := 246, lrValue := 2.298678125671597E+02, bWarn12s := FALSE, bReject13s := FALSE, bReject22s := FALSE),
        (diStep := 247, lrValue := 2.302592494514098E+02, bWarn12s := FALSE, bReject13s := FALSE, bReject22s := FALSE),
        (diStep := 248, lrValue := 2.303004611033681E+02, bWarn12s := FALSE, bReject13s := FALSE, bReject22s := FALSE),
        (diStep := 249, lrValue := 2.295410621479397E+02, bWarn12s := FALSE, bReject13s := FALSE, bReject22s := FALSE),
        (diStep := 250, lrValue := 2.296394750929767E+02, bWarn12s := FALSE, bReject13s := FALSE, bReject22s := FALSE),
        (diStep := 251, lrValue := 2.297358508945258E+02, bWarn12s := FALSE, bReject13s := FALSE, bReject22s := FALSE),
        (diStep := 252, lrValue := 2.299217984946618E+02, bWarn12s := FALSE, bReject13s := FALSE, bReject22s := FALSE),
        (diStep := 253, lrValue := 2.294578388672089E+02, bWarn12s := FALSE, bReject13s := FALSE, bReject22s := FALSE),
        (diStep := 254, lrValue := 2.295892548900854E+02, bWarn12s := FALSE, bReject13s := FALSE, bReject22s := FALSE),
        (diStep := 255, lrValue := 2.297601347464323E+02, bWarn12s := FALSE, bReject13s := FALSE, bReject22s := FALSE),
        (diStep := 256, lrValue := 2.296982505122999E+02, bWarn12s := FALSE, bReject13s := FALSE, bReject22s := FALSE),
        (diStep := 257, lrValue := 2.295729615193367E+02, bWarn12s := FALSE, bReject13s := FALSE, bReject22s := FALSE),
        (diStep := 258, lrValue := 2.296319668314576E+02, bWarn12s := FALSE, bReject13s := FALSE, bReject22s := FALSE),
        (diStep := 259, lrValue := 2.294668115625297E+02, bWarn12s := FALSE, bReject13s := FALSE, bReject22s := FALSE),
        (diStep := 260, lrValue := 2.296908661859453E+02, bWarn12s := FALSE, bReject13s := FALSE, bReject22s := FALSE),
        (diStep := 261, lrValue := 2.297108953449104E+02, bWarn12s := FALSE, bReject13s := FALSE, bReject22s := FALSE),
        (diStep := 262, lrValue := 2.298020877218476E+02, bWarn12s := FALSE, bReject13s := FALSE, bReject22s := FALSE),
        (diStep := 263, lrValue := 2.296836902792228E+02, bWarn12s := FALSE, bReject13s := FALSE, bReject22s := FALSE),
        (diStep := 264, lrValue := 2.298560098055138E+02, bWarn12s := FALSE, bReject13s := FALSE, bReject22s := FALSE),
        (diStep := 265, lrValue := 2.299300144210812E+02, bWarn12s := FALSE, bReject13s := FALSE, bReject22s := FALSE),
        (diStep := 266, lrValue := 2.297755595039245E+02, bWarn12s := FALSE, bReject13s := FALSE, bReject22s := FALSE),
        (diStep := 267, lrValue := 2.298026433801039E+02, bWarn12s := FALSE, bReject13s := FALSE, bReject22s := FALSE),
        (diStep := 268, lrValue := 2.297567883947042E+02, bWarn12s := FALSE, bReject13s := FALSE, bReject22s := FALSE),
        (diStep := 269, lrValue := 2.297575413877743E+02, bWarn12s := FALSE, bReject13s := FALSE, bReject22s := FALSE),
        (diStep := 270, lrValue := 2.296616659484106E+02, bWarn12s := FALSE, bReject13s := FALSE, bReject22s := FALSE),
        (diStep := 271, lrValue := 2.298497051904085E+02, bWarn12s := FALSE, bReject13s := FALSE, bReject22s := FALSE),
        (diStep := 272, lrValue := 2.297927968721062E+02, bWarn12s := FALSE, bReject13s := FALSE, bReject22s := FALSE),
        (diStep := 273, lrValue := 2.301778769710344E+02, bWarn12s := FALSE, bReject13s := FALSE, bReject22s := FALSE),
        (diStep := 274, lrValue := 2.301251916924390E+02, bWarn12s := FALSE, bReject13s := FALSE, bReject22s := FALSE),
        (diStep := 275, lrValue := 2.299933072438744E+02, bWarn12s := FALSE, bReject13s := FALSE, bReject22s := FALSE),
        (diStep := 276, lrValue := 2.299097613406531E+02, bWarn12s := FALSE, bReject13s := FALSE, bReject22s := FALSE),
        (diStep := 277, lrValue := 2.299827547129346E+02, bWarn12s := FALSE, bReject13s := FALSE, bReject22s := FALSE),
        (diStep := 278, lrValue := 2.304589521651602E+02, bWarn12s := FALSE, bReject13s := FALSE, bReject22s := FALSE),
        (diStep := 279, lrValue := 2.303726599951288E+02, bWarn12s := FALSE, bReject13s := FALSE, bReject22s := FALSE),
        (diStep := 280, lrValue := 2.304580352714455E+02, bWarn12s := FALSE, bReject13s := FALSE, bReject22s := FALSE),
        (diStep := 281, lrValue := 2.301154155085727E+02, bWarn12s := FALSE, bReject13s := FALSE, bReject22s := FALSE),
        (diStep := 282, lrValue := 2.305283091889812E+02, bWarn12s := FALSE, bReject13s := FALSE, bReject22s := FALSE),
        (diStep := 283, lrValue := 2.303795450849513E+02, bWarn12s := FALSE, bReject13s := FALSE, bReject22s := FALSE),
        (diStep := 284, lrValue := 2.300553667625987E+02, bWarn12s := FALSE, bReject13s := FALSE, bReject22s := FALSE),
        (diStep := 285, lrValue := 2.301033416478938E+02, bWarn12s := FALSE, bReject13s := FALSE, bReject22s := FALSE),
        (diStep := 286, lrValue := 2.301573457048873E+02, bWarn12s := FALSE, bReject13s := FALSE, bReject22s := FALSE),
        (diStep := 287, lrValue := 2.300508691127785E+02, bWarn12s := FALSE, bReject13s := FALSE, bReject22s := FALSE),
        (diStep := 288, lrValue := 2.299337282370516E+02, bWarn12s := FALSE, bReject13s := FALSE, bReject22s := FALSE),
        (diStep := 289, lrValue := 2.299160610432337E+02, bWarn12s := FALSE, bReject13s := FALSE, bReject22s := FALSE),
        (diStep := 290, lrValue := 2.298535782085829E+02, bWarn12s := FALSE, bReject13s := FALSE, bReject22s := FALSE),
        (diStep := 291, lrValue := 2.298858958705276E+02, bWarn12s := FALSE, bReject13s := FALSE, bReject22s := FALSE),
        (diStep := 292, lrValue := 2.300523485090222E+02, bWarn12s := FALSE, bReject13s := FALSE, bReject22s := FALSE),
        (diStep := 293, lrValue := 2.293845724968881E+02, bWarn12s := TRUE, bReject13s := FALSE, bReject22s := FALSE),
        (diStep := 294, lrValue := 2.297854823900782E+02, bWarn12s := FALSE, bReject13s := FALSE, bReject22s := FALSE),
        (diStep := 295, lrValue := 2.298561685559700E+02, bWarn12s := FALSE, bReject13s := FALSE, bReject22s := FALSE),
        (diStep := 296, lrValue := 2.298627366738675E+02, bWarn12s := FALSE, bReject13s := FALSE, bReject22s := FALSE),
        (diStep := 297, lrValue := 2.297464639181015E+02, bWarn12s := FALSE, bReject13s := FALSE, bReject22s := FALSE),
        (diStep := 298, lrValue := 2.295433810930751E+02, bWarn12s := FALSE, bReject13s := FALSE, bReject22s := FALSE),
        (diStep := 299, lrValue := 2.299039995658953E+02, bWarn12s := FALSE, bReject13s := FALSE, bReject22s := FALSE)
    ];
END_VAR

(* ---- FB_BioPrintPID.st ---- *)
(* =============================================================================
   FB_BioPrintPID — IEC 61131-3 Structured Text port of src/pid_controller.py
   -----------------------------------------------------------------------------
   Parallel PID for a heater zone, called once per task cycle:
     * derivative on measurement (no derivative kick on setpoint steps)
     * first-order filtered derivative, Tf = Kd / (Kp * N)
     * output clamped to [lrOutMin, lrOutMax] (% duty)
     * anti-windup by conditional integration, plus a hard bound on the integrator

   The task cycle time MUST equal lrDt (default T#100MS).
   LREAL is used throughout so that results match the Python reference (IEEE
   double) to ~1e-9 when replaying plc/test_vectors. With REAL, expect
   differences around 1e-3.

   Status: written to match the Python implementation line for line. It has NOT
   been compiled in this repository (no PLC toolchain available here). Verify it with
   tests/FB_BioPrintPID_Test.st (TcUnit) in TwinCAT 3 or CODESYS.
   ============================================================================= *)
FUNCTION_BLOCK FB_BioPrintPID
VAR_INPUT
    lrSetpoint     : LREAL;            (* °C *)
    lrMeasurement  : LREAL;            (* °C, thermocouple *)
    lrKp           : LREAL := 8.0;     (* %/°C *)
    lrKi           : LREAL := 2.5;     (* %/(°C·s) *)
    lrKd           : LREAL := 2.0;     (* %·s/°C *)
    lrDt           : LREAL := 0.1;     (* s, = task cycle time *)
    lrOutMin       : LREAL := 0.0;     (* % *)
    lrOutMax       : LREAL := 100.0;   (* % *)
    lrDerivFilterN : LREAL := 10.0;
    bAntiWindup    : BOOL  := TRUE;
    bReset         : BOOL;             (* clears integrator and derivative memory *)
END_VAR
VAR_OUTPUT
    lrOutput   : LREAL;                (* % duty, clamped *)
    lrPTerm    : LREAL;
    lrITerm    : LREAL;
    lrDTerm    : LREAL;
    bSaturated : BOOL;                 (* TRUE while pushing against a limit *)
END_VAR
VAR
    lrIntegral       : LREAL;
    lrDState         : LREAL;
    lrPrevMeasurement: LREAL;
    bFirstScan       : BOOL := TRUE;
    lrError          : LREAL;
    lrRawD           : LREAL;
    lrTf             : LREAL;
    lrAlpha          : LREAL;
    lrCandidate      : LREAL;
    lrUnclamped      : LREAL;
END_VAR

IF bReset THEN
    lrIntegral := 0.0;
    lrDState   := 0.0;
    bFirstScan := TRUE;
    lrOutput   := 0.0;
    lrPTerm    := 0.0;
    lrITerm    := 0.0;
    lrDTerm    := 0.0;
    bSaturated := FALSE;
    RETURN;
END_IF;

lrError := lrSetpoint - lrMeasurement;

(* --- Derivative on measurement, low-pass filtered ------------------------- *)
IF bFirstScan THEN
    lrRawD := 0.0;
    bFirstScan := FALSE;
ELSE
    lrRawD := -(lrMeasurement - lrPrevMeasurement) / lrDt;
END_IF;
lrPrevMeasurement := lrMeasurement;

IF lrKp > 0.0 AND lrDerivFilterN > 0.0 THEN
    lrTf := lrKd / (lrKp * lrDerivFilterN);
ELSE
    lrTf := 0.0;
END_IF;
IF lrTf > 0.0 THEN
    lrAlpha := lrDt / (lrTf + lrDt);
ELSE
    lrAlpha := 1.0;
END_IF;
lrDState := lrDState + lrAlpha * (lrRawD - lrDState);

lrPTerm := lrKp * lrError;
lrDTerm := lrKd * lrDState;

(* --- Integral with conditional integration (anti-windup) ------------------ *)
lrCandidate := lrIntegral + lrKi * lrError * lrDt;
lrUnclamped := lrPTerm + lrCandidate + lrDTerm;
bSaturated  := (lrUnclamped > lrOutMax AND lrError > 0.0)
            OR (lrUnclamped < lrOutMin AND lrError < 0.0);

IF NOT (bAntiWindup AND bSaturated) THEN
    lrIntegral := lrCandidate;
END_IF;
IF bAntiWindup THEN
    (* Hard bound as a second line of defence against numerical drift *)
    lrIntegral := LIMIT(lrOutMin, lrIntegral, lrOutMax);
END_IF;

lrITerm  := lrIntegral;
lrOutput := LIMIT(lrOutMin, lrPTerm + lrIntegral + lrDTerm, lrOutMax);
END_FUNCTION_BLOCK

(* ---- FB_WestgardMonitor.st ---- *)
(* =============================================================================
   FB_WestgardMonitor — IEC 61131-3 Structured Text port of src/westgard_validator.py
   -----------------------------------------------------------------------------
   Clinical Westgard multirule on one process variable, called once per sample:
     Phase 1  collect iBaselineLength samples from diBaselineStart, then fix the SD
              (sample SD, n-1) with a floor of lrMinSd
     Phase 2  judge each later sample against lrTarget ± k·SD
                1-2s  warning   |z| > 2
                1-3s  reject    |z| > 3
                2-2s  reject    two consecutive |z| > 2 on the same side
   bRunRejected latches until bReset, like a rejected analytical run in a lab.

   Not ported: rolling mean / SD / CV% (dashboard statistics only).
   Status: NOT compiled in this repository. Verify with tests/FB_WestgardMonitor_Test.st.
   ============================================================================= *)
FUNCTION_BLOCK FB_WestgardMonitor
VAR_INPUT
    lrValue          : LREAL;          (* sample, e.g. barrel temperature °C *)
    lrTarget         : LREAL := 230.0; (* assigned value, i.e. the setpoint *)
    diStep           : DINT;           (* sample index, starting at 0 *)
    diBaselineStart  : DINT := 80;
    iBaselineLength  : INT  := 40;     (* 10 .. MAX_BASELINE *)
    lrMinSd          : LREAL := 0.05;
    bReset           : BOOL;
END_VAR
VAR_OUTPUT
    bArmed        : BOOL;              (* baseline fixed, rules active *)
    lrBaselineSd  : LREAL;
    lrZ           : LREAL;
    bWarn12s      : BOOL;              (* this sample *)
    bReject13s    : BOOL;              (* this sample *)
    bReject22s    : BOOL;              (* this sample *)
    bRunRejected  : BOOL;              (* latched *)
    bConfigError  : BOOL;
END_VAR
VAR CONSTANT
    MAX_BASELINE : INT := 200;
END_VAR
VAR
    alrBaseline : ARRAY[1..200] OF LREAL;
    iCount      : INT;
    i           : INT;
    lrSum       : LREAL;
    lrMean      : LREAL;
    lrSq        : LREAL;
    lrPrevZ     : LREAL;
    bHavePrev   : BOOL;
END_VAR

IF bReset THEN
    iCount := 0; bArmed := FALSE; bHavePrev := FALSE; bRunRejected := FALSE;
    lrBaselineSd := 0.0; lrZ := 0.0;
END_IF;

bWarn12s := FALSE;
bReject13s := FALSE;
bReject22s := FALSE;
bConfigError := (iBaselineLength < 10) OR (iBaselineLength > MAX_BASELINE);
IF bConfigError THEN
    RETURN;
END_IF;

(* --- Phase 1: baseline window ---------------------------------------------- *)
IF diStep >= diBaselineStart AND diStep < diBaselineStart + INT_TO_DINT(iBaselineLength) THEN
    iCount := iCount + 1;
    alrBaseline[iCount] := lrValue;
    IF iCount = iBaselineLength THEN
        lrSum := 0.0;
        FOR i := 1 TO iCount DO
            lrSum := lrSum + alrBaseline[i];
        END_FOR;
        lrMean := lrSum / INT_TO_LREAL(iCount);
        lrSq := 0.0;
        FOR i := 1 TO iCount DO
            lrSq := lrSq + (alrBaseline[i] - lrMean) * (alrBaseline[i] - lrMean);
        END_FOR;
        lrBaselineSd := MAX(SQRT(lrSq / INT_TO_LREAL(iCount - 1)), lrMinSd);
        bArmed := TRUE;
    END_IF;
    RETURN;
END_IF;

IF NOT bArmed THEN
    RETURN;
END_IF;

(* --- Phase 2: Westgard rules against target and fixed SD ------------------- *)
lrZ := (lrValue - lrTarget) / lrBaselineSd;

IF ABS(lrZ) > 3.0 THEN
    bReject13s := TRUE;
ELSIF ABS(lrZ) > 2.0 THEN
    bWarn12s := TRUE;
END_IF;

IF bHavePrev AND ABS(lrZ) > 2.0 AND ABS(lrPrevZ) > 2.0
   AND ((lrZ > 0.0) = (lrPrevZ > 0.0)) THEN
    bReject22s := TRUE;
END_IF;

lrPrevZ := lrZ;
bHavePrev := TRUE;
bRunRejected := bRunRejected OR bReject13s OR bReject22s;
END_FUNCTION_BLOCK
